(* IEC 61131-3 sources: plc-vscode/tests/st/test-ready/trust-platform/libraries/oscat/oop/src, 12 files *)

(* ---- component_types.st ---- *)
TYPE ComponentStatus :
STRUCT
    Ready : BOOL;
    Error : BOOL;
    ErrorId : WORD;
    Status : BYTE;
END_STRUCT
END_TYPE

TYPE RealRange :
STRUCT
    Low : REAL;
    High : REAL;
END_STRUCT
END_TYPE

TYPE PidGains :
STRUCT
    Kp : REAL := 1.0;
    Tn : REAL := 1.0;
    Tv : REAL := 1.0;
END_STRUCT
END_TYPE

TYPE PiGains :
STRUCT
    Kp : REAL := 1.0;
    Ki : REAL := 1.0;
END_STRUCT
END_TYPE

TYPE SunPosition :
STRUCT
    Azimuth : REAL;
    Elevation : REAL;
    RefractedElevation : REAL;
END_STRUCT
END_TYPE

TYPE SunTimes :
STRUCT
    SolarNoon : TOD;
    Sunrise : TOD;
    Sunset : TOD;
    Declination : REAL;
END_STRUCT
END_TYPE

TYPE BarGraphSnapshot :
STRUCT
    Low : BOOL;
    Q1 : BOOL;
    Q2 : BOOL;
    Q3 : BOOL;
    Q4 : BOOL;
    Q5 : BOOL;
    Q6 : BOOL;
    High : BOOL;
    Alarm : BOOL;
    Status : BYTE;
END_STRUCT
END_TYPE

VAR_GLOBAL CONSTANT
    ComponentErrorNone : WORD := WORD#16#0000;
    ComponentErrorInvalidConfiguration : WORD := WORD#16#1000;
    ComponentErrorNotReady : WORD := WORD#16#1001;
    ComponentErrorQueueFull : WORD := WORD#16#1002;
    ComponentErrorQueueEmpty : WORD := WORD#16#1003;

    DefaultPidKp : REAL := REAL#1.0;
    DefaultPidTn : REAL := REAL#1.0;
    DefaultPidTv : REAL := REAL#1.0;
    DefaultPidLowLimit : REAL := REAL#-1000.0;
    DefaultPidHighLimit : REAL := REAL#1000.0;
    DefaultPidSupervisionBand : REAL := REAL#0.0;
    DefaultPidOffset : REAL := REAL#0.0;

    DefaultPt1Gain : REAL := REAL#1.0;
    DefaultPt1TimeConstant : TIME := T#1s;
    DefaultPulseHighTime : TIME := T#1s;
    DefaultPulseLowTime : TIME := T#1s;
    DefaultCalendarOffsetMinutes : INT := INT#0;
    MaxDwordFifo16Capacity : UINT := UINT#16;
    MaxDwordStack16Capacity : UINT := UINT#16;
    MaxDwordFifo32Capacity : UINT := UINT#32;
    MaxDwordStack32Capacity : UINT := UINT#32;
END_VAR

(* ---- component_interfaces.st ---- *)
INTERFACE IComponent
    PROPERTY Ready : BOOL
    GET
    END_GET
    END_PROPERTY

    PROPERTY Error : BOOL
    GET
    END_GET
    END_PROPERTY

    PROPERTY ErrorId : WORD
    GET
    END_GET
    END_PROPERTY

    PROPERTY Status : BYTE
    GET
    END_GET
    END_PROPERTY

    METHOD Initialize
    END_METHOD

    METHOD Reset
    END_METHOD

    METHOD ClearError
    END_METHOD

    METHOD Snapshot : ComponentStatus
    END_METHOD
END_INTERFACE

INTERFACE IAutomationContext EXTENDS IComponent
    PROPERTY ConstantsLoaded : BOOL
    GET
    END_GET
    END_PROPERTY

    PROPERTY Version : DWORD
    GET
    END_GET
    END_PROPERTY

    PROPERTY Math : CONSTANTS_MATH
    GET
    END_GET
    END_PROPERTY

    PROPERTY Pi2 : REAL
    GET
    END_GET
    END_PROPERTY

    PROPERTY Phys : CONSTANTS_PHYS
    GET
    END_GET
    END_PROPERTY

    PROPERTY LanguageValues : CONSTANTS_LANGUAGE
    GET
    END_GET
    END_PROPERTY

    PROPERTY DefaultLanguage : INT
    GET
    END_GET
    END_PROPERTY

    METHOD LoadConstants : BOOL
    END_METHOD

    METHOD SetDefaultLanguage
    VAR_INPUT
        LanguageIndex : INT;
    END_VAR
    END_METHOD

    METHOD DirectionName : STRING[3]
    VAR_INPUT
        Degrees : REAL;
    END_VAR
    END_METHOD

    METHOD DirectionDegrees : INT
    VAR_INPUT
        Name : STRING[3];
    END_VAR
    END_METHOD
END_INTERFACE

INTERFACE IUnitConverter EXTENDS IComponent
    METHOD KelvinFromCelsius : REAL
    VAR_INPUT
        Celsius : REAL;
    END_VAR
    END_METHOD

    METHOD FahrenheitFromCelsius : REAL
    VAR_INPUT
        Celsius : REAL;
    END_VAR
    END_METHOD

    METHOD CelsiusFromKelvin : REAL
    VAR_INPUT
        Kelvin : REAL;
    END_VAR
    END_METHOD

    METHOD CelsiusFromFahrenheit : REAL
    VAR_INPUT
        Fahrenheit : REAL;
    END_VAR
    END_METHOD

    METHOD MetersPerSecondFromKilometersPerHour : REAL
    VAR_INPUT
        Kmh : REAL;
    END_VAR
    END_METHOD

    METHOD KilometersPerHourFromMetersPerSecond : REAL
    VAR_INPUT
        Mps : REAL;
    END_VAR
    END_METHOD

    METHOD BeaufortFromMetersPerSecond : INT
    VAR_INPUT
        Mps : REAL;
    END_VAR
    END_METHOD

    METHOD AngularFrequencyFromHertz : REAL
    VAR_INPUT
        Frequency : REAL;
    END_VAR
    END_METHOD

    METHOD HertzFromAngularFrequency : REAL
    VAR_INPUT
        AngularFrequency : REAL;
    END_VAR
    END_METHOD

    METHOD PeriodFromHertz : TIME
    VAR_INPUT
        Frequency : REAL;
    END_VAR
    END_METHOD

    METHOD HertzFromPeriod : REAL
    VAR_INPUT
        Period : TIME;
    END_VAR
    END_METHOD

    METHOD WattHoursFromJoules : REAL
    VAR_INPUT
        Joule : REAL;
    END_VAR
    END_METHOD

    METHOD JoulesFromWattHours : REAL
    VAR_INPUT
        WattHour : REAL;
    END_VAR
    END_METHOD

    METHOD JoulesFromCalories : REAL
    VAR_INPUT
        Calorie : REAL;
    END_VAR
    END_METHOD

    METHOD CaloriesFromJoules : REAL
    VAR_INPUT
        Joule : REAL;
    END_VAR
    END_METHOD
END_INTERFACE

INTERFACE IPt1Filter EXTENDS IComponent
    PROPERTY Output : REAL
    GET
    END_GET
    END_PROPERTY

    PROPERTY TimeConstant : TIME
    GET
    END_GET
    END_PROPERTY

    PROPERTY Gain : REAL
    GET
    END_GET
    END_PROPERTY

    METHOD Configure
    VAR_INPUT
        TimeConstant : TIME;
        Gain : REAL;
    END_VAR
    END_METHOD

    METHOD Update : REAL
    VAR_INPUT
        Sample : REAL;
    END_VAR
    END_METHOD
END_INTERFACE

INTERFACE IClosedLoopController EXTENDS IComponent
    PROPERTY Actual : REAL
    GET
    END_GET
    END_PROPERTY

    PROPERTY TargetValue : REAL
    GET
    END_GET
    END_PROPERTY

    PROPERTY Output : REAL
    GET
    END_GET
    END_PROPERTY

    PROPERTY ControlError : REAL
    GET
    END_GET
    END_PROPERTY

    PROPERTY Limited : BOOL
    GET
    END_GET
    END_PROPERTY

    METHOD Update : REAL
    VAR_INPUT
        Actual : REAL;
        Target : REAL;
    END_VAR
    END_METHOD
END_INTERFACE

INTERFACE IPidController EXTENDS IClosedLoopController
    PROPERTY SupervisionBand : REAL
    GET
    END_GET
    END_PROPERTY

    PROPERTY Manual : BOOL
    GET
    END_GET
    END_PROPERTY

    PROPERTY ManualInput : REAL
    GET
    END_GET
    END_PROPERTY

    PROPERTY Offset : REAL
    GET
    END_GET
    END_PROPERTY

    PROPERTY LowLimit : REAL
    GET
    END_GET
    END_PROPERTY

    PROPERTY HighLimit : REAL
    GET
    END_GET
    END_PROPERTY

    PROPERTY Kp : REAL
    GET
    END_GET
    END_PROPERTY

    PROPERTY Tn : REAL
    GET
    END_GET
    END_PROPERTY

    PROPERTY Tv : REAL
    GET
    END_GET
    END_PROPERTY

    METHOD SetKp
    VAR_INPUT
        Kp : REAL;
    END_VAR
    END_METHOD

    METHOD SetIntegralTime
    VAR_INPUT
        Tn : REAL;
    END_VAR
    END_METHOD

    METHOD SetDerivativeTime
    VAR_INPUT
        Tv : REAL;
    END_VAR
    END_METHOD

    METHOD SetSupervisionBand
    VAR_INPUT
        SupervisionBand : REAL;
    END_VAR
    END_METHOD

    METHOD SetOffset
    VAR_INPUT
        Offset : REAL;
    END_VAR
    END_METHOD

    METHOD SetLimits
    VAR_INPUT
        Limits : RealRange;
    END_VAR
    END_METHOD

    METHOD SetManual
    VAR_INPUT
        Manual : BOOL;
        ManualInput : REAL;
    END_VAR
    END_METHOD

    METHOD ApplyGains
    VAR_INPUT
        Gains : PidGains;
    END_VAR
    END_METHOD

    METHOD Configure
    VAR_INPUT
        Gains : PidGains;
        Limits : RealRange;
        SupervisionBand : REAL;
        Offset : REAL;
    END_VAR
    END_METHOD

END_INTERFACE

INTERFACE IHysteresisSwitch EXTENDS IComponent
    PROPERTY MeasuredValue : REAL
    GET
    END_GET
    END_PROPERTY

    PROPERTY LowLimit : REAL
    GET
    END_GET
    END_PROPERTY

    PROPERTY HighLimit : REAL
    GET
    END_GET
    END_PROPERTY

    PROPERTY Q : BOOL
    GET
    END_GET
    END_PROPERTY

    PROPERTY Window : BOOL
    GET
    END_GET
    END_PROPERTY

    METHOD SetLimits
    VAR_INPUT
        Limits : RealRange;
    END_VAR
    END_METHOD

    METHOD Update : BOOL
    VAR_INPUT
        MeasuredValue : REAL;
    END_VAR
    END_METHOD
END_INTERFACE

INTERFACE IPulseGenerator EXTENDS IComponent
    PROPERTY Enabled : BOOL
    GET
    END_GET
    END_PROPERTY

    PROPERTY Output : BOOL
    GET
    END_GET
    END_PROPERTY

    PROPERTY HighTime : TIME
    GET
    END_GET
    END_PROPERTY

    PROPERTY LowTime : TIME
    GET
    END_GET
    END_PROPERTY

    METHOD Configure
    VAR_INPUT
        HighTime : TIME;
        LowTime : TIME;
    END_VAR
    END_METHOD

    METHOD SetEnabled
    VAR_INPUT
        Enabled : BOOL;
    END_VAR
    END_METHOD

    METHOD Update : BOOL
    END_METHOD
END_INTERFACE

INTERFACE IDwordQueue EXTENDS IComponent
    PROPERTY Empty : BOOL
    GET
    END_GET
    END_PROPERTY

    PROPERTY Full : BOOL
    GET
    END_GET
    END_PROPERTY

    PROPERTY Value : DWORD
    GET
    END_GET
    END_PROPERTY

    PROPERTY Capacity : UINT
    GET
    END_GET
    END_PROPERTY

    METHOD Push : BOOL
    VAR_INPUT
        Value : DWORD;
    END_VAR
    END_METHOD

    METHOD TryPop : BOOL
    END_METHOD
END_INTERFACE

INTERFACE IDwordStack EXTENDS IComponent
    PROPERTY Empty : BOOL
    GET
    END_GET
    END_PROPERTY

    PROPERTY Full : BOOL
    GET
    END_GET
    END_PROPERTY

    PROPERTY Value : DWORD
    GET
    END_GET
    END_PROPERTY

    PROPERTY Capacity : UINT
    GET
    END_GET
    END_PROPERTY

    METHOD Push : BOOL
    VAR_INPUT
        Value : DWORD;
    END_VAR
    END_METHOD

    METHOD TryPop : BOOL
    END_METHOD
END_INTERFACE

INTERFACE ICalendarClock EXTENDS IComponent
    PROPERTY Utc : DT
    GET
    END_GET
    END_PROPERTY

    PROPERTY LocalDateTime : DT
    GET
    END_GET
    END_PROPERTY

    PROPERTY LocalDate : DATE
    GET
    END_GET
    END_PROPERTY

    PROPERTY LocalTimeOfDay : TOD
    GET
    END_GET
    END_PROPERTY

    PROPERTY Year : INT
    GET
    END_GET
    END_PROPERTY

    PROPERTY Month : INT
    GET
    END_GET
    END_PROPERTY

    PROPERTY Day : INT
    GET
    END_GET
    END_PROPERTY

    PROPERTY Weekday : INT
    GET
    END_GET
    END_PROPERTY

    PROPERTY OffsetMinutes : INT
    GET
    END_GET
    END_PROPERTY

    PROPERTY DstEnabled : BOOL
    GET
    END_GET
    END_PROPERTY

    PROPERTY DstOn : BOOL
    GET
    END_GET
    END_PROPERTY

    PROPERTY LanguageIndex : INT
    GET
    END_GET
    END_PROPERTY

    PROPERTY Longitude : REAL
    GET
    END_GET
    END_PROPERTY

    PROPERTY Latitude : REAL
    GET
    END_GET
    END_PROPERTY

    PROPERTY Sunrise : TOD
    GET
    END_GET
    END_PROPERTY

    PROPERTY Sunset : TOD
    GET
    END_GET
    END_PROPERTY

    PROPERTY SolarNoon : TOD
    GET
    END_GET
    END_PROPERTY

    PROPERTY SolarElevation : REAL
    GET
    END_GET
    END_PROPERTY

    PROPERTY SolarHorizontalProjection : REAL
    GET
    END_GET
    END_PROPERTY

    PROPERTY SolarVerticalProjection : REAL
    GET
    END_GET
    END_PROPERTY

    PROPERTY Night : BOOL
    GET
    END_GET
    END_PROPERTY

    PROPERTY Holiday : BOOL
    GET
    END_GET
    END_PROPERTY

    PROPERTY HolidayName : STRING[30]
    GET
    END_GET
    END_PROPERTY

    PROPERTY WorkWeek : INT
    GET
    END_GET
    END_PROPERTY

    METHOD Configure
    VAR_INPUT
        LocationLatitude : REAL;
        LocationLongitude : REAL;
        OffsetMinutes : INT;
        DstEnabled : BOOL;
        LanguageIndex : INT;
    END_VAR
    END_METHOD

    METHOD Update
    VAR_INPUT
        Utc : DT;
    END_VAR
    END_METHOD

    METHOD CalculateSunPosition : SunPosition
    VAR_INPUT
        Utc : DT;
        Latitude : REAL;
        Longitude : REAL;
    END_VAR
    END_METHOD

    METHOD CalculateSunTime : SunTimes
    VAR_INPUT
        UtcDate : DATE;
        Latitude : REAL;
        Longitude : REAL;
        Horizon : REAL;
    END_VAR
    END_METHOD
END_INTERFACE

(* ---- automation_context.st ---- *)
FUNCTION_BLOCK AutomationContext IMPLEMENTS IAutomationContext
VAR
    ReadyValue : BOOL;
    ErrorValue : BOOL;
    ErrorIdValue : WORD;
    StatusValue : BYTE;
    ConstantsLoadedValue : BOOL;
END_VAR

METHOD PUBLIC Initialize
ApplyConstantsLoadResult(Loaded := OSCAT_BASIC_Constants());
END_METHOD

METHOD PUBLIC Reset
ClearError();
ConstantsLoadedValue := FALSE;
END_METHOD

METHOD PUBLIC ClearError
ErrorValue := FALSE;
ErrorIdValue := ComponentErrorNone;
StatusValue := BYTE#0;
END_METHOD

METHOD PUBLIC Snapshot : ComponentStatus
VAR
    Result : ComponentStatus;
END_VAR
Result.Ready := ReadyValue;
Result.Error := ErrorValue;
Result.ErrorId := ErrorIdValue;
Result.Status := StatusValue;
Snapshot := Result;
END_METHOD

METHOD PUBLIC LoadConstants : BOOL
LoadConstants := OSCAT_BASIC_Constants();
ApplyConstantsLoadResult(Loaded := LoadConstants);
END_METHOD

METHOD PRIVATE ApplyConstantsLoadResult
VAR_INPUT
    Loaded : BOOL;
END_VAR
ConstantsLoadedValue := Loaded;
ReadyValue := Loaded;
IF Loaded THEN
    ClearError();
ELSE
    ErrorValue := TRUE;
    ErrorIdValue := ComponentErrorNotReady;
    StatusValue := BYTE#1;
END_IF;
END_METHOD

METHOD PUBLIC SetDefaultLanguage
VAR_INPUT
    LanguageIndex : INT;
END_VAR
IF NOT ConstantsLoadedValue AND NOT LoadConstants() THEN
    ErrorValue := TRUE;
    ErrorIdValue := ComponentErrorNotReady;
    StatusValue := BYTE#1;
ELSIF LanguageIndex >= INT#1 AND LanguageIndex <= LANGUAGE.LMAX THEN
    LANGUAGE.DEFAULT := LanguageIndex;
    ClearError();
ELSE
    ErrorValue := TRUE;
    ErrorIdValue := ComponentErrorInvalidConfiguration;
    StatusValue := BYTE#1;
END_IF;
END_METHOD

METHOD PUBLIC DirectionName : STRING[3]
VAR_INPUT
    Degrees : REAL;
END_VAR
IF NOT ConstantsLoadedValue AND NOT LoadConstants() THEN
    DirectionName := '';
ELSE
    DirectionName := DEG_TO_DIR(DEG := REAL_TO_INT(Degrees), N := INT#4, L := LANGUAGE.DEFAULT);
END_IF;
END_METHOD

METHOD PUBLIC DirectionDegrees : INT
VAR_INPUT
    Name : STRING[3];
END_VAR
IF NOT ConstantsLoadedValue AND NOT LoadConstants() THEN
    DirectionDegrees := INT#0;
ELSE
    DirectionDegrees := DIR_TO_DEG(DIR := Name, L := LANGUAGE.DEFAULT);
END_IF;
END_METHOD

PUBLIC PROPERTY Ready : BOOL
GET
    Ready := ReadyValue;
END_GET
END_PROPERTY

PUBLIC PROPERTY Error : BOOL
GET
    Error := ErrorValue;
END_GET
END_PROPERTY

PUBLIC PROPERTY ErrorId : WORD
GET
    ErrorId := ErrorIdValue;
END_GET
END_PROPERTY

PUBLIC PROPERTY Status : BYTE
GET
    Status := StatusValue;
END_GET
END_PROPERTY

PUBLIC PROPERTY ConstantsLoaded : BOOL
GET
    ConstantsLoaded := ConstantsLoadedValue OR g_oscat_constants_loaded;
END_GET
END_PROPERTY

PUBLIC PROPERTY Version : DWORD
GET
    Version := OSCAT_VERSION(IN := FALSE);
END_GET
END_PROPERTY

PUBLIC PROPERTY Math : CONSTANTS_MATH
GET
    Math := MATH;
END_GET
END_PROPERTY

PUBLIC PROPERTY Pi2 : REAL
GET
    Pi2 := MATH.PI2;
END_GET
END_PROPERTY

PUBLIC PROPERTY Phys : CONSTANTS_PHYS
GET
    Phys := PHYS;
END_GET
END_PROPERTY

PUBLIC PROPERTY LanguageValues : CONSTANTS_LANGUAGE
GET
    LanguageValues := LANGUAGE;
END_GET
END_PROPERTY

PUBLIC PROPERTY DefaultLanguage : INT
GET
    DefaultLanguage := LANGUAGE.DEFAULT;
END_GET
END_PROPERTY
END_FUNCTION_BLOCK

(* ---- calendar.st ---- *)
FUNCTION_BLOCK CalendarClock IMPLEMENTS ICalendarClock
VAR
    ReadyValue : BOOL;
    ErrorValue : BOOL;
    ErrorIdValue : WORD;
    StatusValue : BYTE;
    CalendarData : CALENDAR;
    Holidays : ARRAY[0..29] OF HOLIDAY_DATA;
    CalendarFb : CALENDAR_CALC;
    SunPositionFb : SUN_POS;
    SunTimeFb : SUN_TIME;
END_VAR

METHOD PUBLIC Initialize
ReadyValue := TRUE;
OSCAT_BASIC_Constants();
CalendarData.OFFSET := DefaultCalendarOffsetMinutes;
CalendarData.LANGUAGE := LANGUAGE.DEFAULT;
ClearError();
END_METHOD

METHOD PUBLIC Reset
ClearError();
END_METHOD

METHOD PUBLIC ClearError
ErrorValue := FALSE;
ErrorIdValue := ComponentErrorNone;
StatusValue := BYTE#0;
END_METHOD

METHOD PUBLIC Snapshot : ComponentStatus
VAR
    Result : ComponentStatus;
END_VAR
Result.Ready := ReadyValue;
Result.Error := ErrorValue;
Result.ErrorId := ErrorIdValue;
Result.Status := StatusValue;
Snapshot := Result;
END_METHOD

METHOD PUBLIC Configure
VAR_INPUT
    LocationLatitude : REAL;
    LocationLongitude : REAL;
    OffsetMinutes : INT;
    DstEnabled : BOOL;
    LanguageIndex : INT;
END_VAR
IF NOT ReadyValue THEN
    Initialize();
END_IF;
CalendarData.LATITUDE := LocationLatitude;
CalendarData.LONGITUDE := LocationLongitude;
CalendarData.OFFSET := OffsetMinutes;
CalendarData.DST_EN := DstEnabled;
CalendarData.LANGUAGE := LanguageIndex;
ClearError();
END_METHOD

METHOD PUBLIC Update
VAR_INPUT
    Utc : DT;
END_VAR
IF NOT ReadyValue THEN
    Initialize();
END_IF;
CalendarData.UTC := Utc;
CalendarFb(SPE := TRUE, H := REAL#-0.8333333, XCAL := CalendarData, HOLIDAYS := Holidays);
END_METHOD

METHOD PUBLIC CalculateSunPosition : SunPosition
VAR_INPUT
    Utc : DT;
    Latitude : REAL;
    Longitude : REAL;
END_VAR
VAR
    Result : SunPosition;
END_VAR
OSCAT_BASIC_Constants();
SunPositionFb(LATITUDE := Latitude, LONGITUDE := Longitude, UTC := Utc);
Result.Azimuth := SunPositionFb.B;
Result.Elevation := SunPositionFb.H;
Result.RefractedElevation := SunPositionFb.HR;
CalculateSunPosition := Result;
END_METHOD

METHOD PUBLIC CalculateSunTime : SunTimes
VAR_INPUT
    UtcDate : DATE;
    Latitude : REAL;
    Longitude : REAL;
    Horizon : REAL;
END_VAR
VAR
    Result : SunTimes;
END_VAR
OSCAT_BASIC_Constants();
SunTimeFb(LATITUDE := Latitude, LONGITUDE := Longitude, UTC := UtcDate, H := Horizon);
Result.SolarNoon := SunTimeFb.MIDDAY;
Result.Sunrise := SunTimeFb.SUN_RISE;
Result.Sunset := SunTimeFb.SUN_SET;
Result.Declination := SunTimeFb.SUN_DECLINATION;
CalculateSunTime := Result;
END_METHOD

PUBLIC PROPERTY Ready : BOOL
GET
    Ready := ReadyValue;
END_GET
END_PROPERTY

PUBLIC PROPERTY Error : BOOL
GET
    Error := ErrorValue;
END_GET
END_PROPERTY

PUBLIC PROPERTY ErrorId : WORD
GET
    ErrorId := ErrorIdValue;
END_GET
END_PROPERTY

PUBLIC PROPERTY Status : BYTE
GET
    Status := StatusValue;
END_GET
END_PROPERTY

PUBLIC PROPERTY Utc : DT
GET
    Utc := CalendarData.UTC;
END_GET
END_PROPERTY

PUBLIC PROPERTY LocalDateTime : DT
GET
    LocalDateTime := CalendarData.LOCAL_DT;
END_GET
END_PROPERTY

PUBLIC PROPERTY LocalDate : DATE
GET
    LocalDate := CalendarData.LOCAL_DATE;
END_GET
END_PROPERTY

PUBLIC PROPERTY LocalTimeOfDay : TOD
GET
    LocalTimeOfDay := CalendarData.LOCAL_TOD;
END_GET
END_PROPERTY

PUBLIC PROPERTY Year : INT
GET
    Year := CalendarData.YEAR;
END_GET
END_PROPERTY

PUBLIC PROPERTY Month : INT
GET
    Month := CalendarData.MONTH;
END_GET
END_PROPERTY

PUBLIC PROPERTY Day : INT
GET
    Day := CalendarData.DAY;
END_GET
END_PROPERTY

PUBLIC PROPERTY Weekday : INT
GET
    Weekday := CalendarData.WEEKDAY;
END_GET
END_PROPERTY

PUBLIC PROPERTY OffsetMinutes : INT
GET
    OffsetMinutes := CalendarData.OFFSET;
END_GET
END_PROPERTY

PUBLIC PROPERTY DstEnabled : BOOL
GET
    DstEnabled := CalendarData.DST_EN;
END_GET
END_PROPERTY

PUBLIC PROPERTY DstOn : BOOL
GET
    DstOn := CalendarData.DST_ON;
END_GET
END_PROPERTY

PUBLIC PROPERTY LanguageIndex : INT
GET
    LanguageIndex := CalendarData.LANGUAGE;
END_GET
END_PROPERTY

PUBLIC PROPERTY Longitude : REAL
GET
    Longitude := CalendarData.LONGITUDE;
END_GET
END_PROPERTY

PUBLIC PROPERTY Latitude : REAL
GET
    Latitude := CalendarData.LATITUDE;
END_GET
END_PROPERTY

PUBLIC PROPERTY Sunrise : TOD
GET
    Sunrise := CalendarData.SUN_RISE;
END_GET
END_PROPERTY

PUBLIC PROPERTY Sunset : TOD
GET
    Sunset := CalendarData.SUN_SET;
END_GET
END_PROPERTY

PUBLIC PROPERTY SolarNoon : TOD
GET
    SolarNoon := CalendarData.SUN_MIDDAY;
END_GET
END_PROPERTY

PUBLIC PROPERTY SolarElevation : REAL
GET
    (* OSCAT classic keeps the historical SUN_HEIGTH spelling. *)
    SolarElevation := CalendarData.SUN_HEIGTH;
END_GET
END_PROPERTY

PUBLIC PROPERTY SolarHorizontalProjection : REAL
GET
    SolarHorizontalProjection := CalendarData.SUN_HOR;
END_GET
END_PROPERTY

PUBLIC PROPERTY SolarVerticalProjection : REAL
GET
    SolarVerticalProjection := CalendarData.SUN_VER;
END_GET
END_PROPERTY

PUBLIC PROPERTY Night : BOOL
GET
    Night := CalendarData.NIGHT;
END_GET
END_PROPERTY

PUBLIC PROPERTY Holiday : BOOL
GET
    Holiday := CalendarData.HOLIDAY;
END_GET
END_PROPERTY

PUBLIC PROPERTY HolidayName : STRING[30]
GET
    HolidayName := CalendarData.HOLY_NAME;
END_GET
END_PROPERTY

PUBLIC PROPERTY WorkWeek : INT
GET
    WorkWeek := CalendarData.WORK_WEEK;
END_GET
END_PROPERTY
END_FUNCTION_BLOCK

FUNCTION_BLOCK HolidayCalendar IMPLEMENTS IComponent
VAR
    ReadyValue : BOOL;
    ErrorValue : BOOL;
    ErrorIdValue : WORD;
    StatusValue : BYTE;
    HolidayValue : BOOL;
    NameValue : STRING[30];
    LanguageIndexValue : INT := INT#1;
    FridayAsHolidayValue : BOOL;
    SaturdayAsHolidayValue : BOOL;
    SundayAsHolidayValue : BOOL;
    Holidays : ARRAY[0..29] OF HOLIDAY_DATA;
    HolidayFb : HOLIDAY;
END_VAR

METHOD PUBLIC Initialize
ReadyValue := TRUE;
OSCAT_BASIC_Constants();
ClearError();
END_METHOD

METHOD PUBLIC Reset
HolidayValue := FALSE;
NameValue := '';
ClearError();
END_METHOD

METHOD PUBLIC ClearError
ErrorValue := FALSE;
ErrorIdValue := ComponentErrorNone;
StatusValue := BYTE#0;
END_METHOD

METHOD PUBLIC Snapshot : ComponentStatus
VAR
    Result : ComponentStatus;
END_VAR
Result.Ready := ReadyValue;
Result.Error := ErrorValue;
Result.ErrorId := ErrorIdValue;
Result.Status := StatusValue;
Snapshot := Result;
END_METHOD

METHOD PUBLIC Configure
VAR_INPUT
    LanguageIndex : INT;
    FridayAsHoliday : BOOL;
    SaturdayAsHoliday : BOOL;
    SundayAsHoliday : BOOL;
END_VAR
LanguageIndexValue := LanguageIndex;
FridayAsHolidayValue := FridayAsHoliday;
SaturdayAsHolidayValue := SaturdayAsHoliday;
SundayAsHolidayValue := SundayAsHoliday;
ClearError();
END_METHOD

METHOD PUBLIC SetHoliday
VAR_INPUT
    Index : INT;
    Month : SINT;
    Day : SINT;
    Use : SINT;
    Name : STRING[30];
END_VAR
IF Index < INT#0 OR Index > INT#29 THEN
    ErrorValue := TRUE;
    ErrorIdValue := ComponentErrorInvalidConfiguration;
    StatusValue := BYTE#1;
ELSE
    Holidays[Index].MONTH := Month;
    Holidays[Index].DAY := Day;
    Holidays[Index].USE := Use;
    Holidays[Index].NAME := Name;
    ClearError();
END_IF;
END_METHOD

METHOD PUBLIC Update : BOOL
VAR_INPUT
    DateIn : DATE;
END_VAR
HolidayFb(
    DATE_IN := DateIn,
    LANGU := LanguageIndexValue,
    FRIDAY := FridayAsHolidayValue,
    SATURDAY := SaturdayAsHolidayValue,
    SUNDAY := SundayAsHolidayValue,
    HOLIDAYS := Holidays
);
HolidayValue := HolidayFb.Y;
NameValue := HolidayFb.NAME;
Update := HolidayValue;
END_METHOD

PUBLIC PROPERTY Ready : BOOL
GET
    Ready := ReadyValue;
END_GET
END_PROPERTY

PUBLIC PROPERTY Error : BOOL
GET
    Error := ErrorValue;
END_GET
END_PROPERTY

PUBLIC PROPERTY ErrorId : WORD
GET
    ErrorId := ErrorIdValue;
END_GET
END_PROPERTY

PUBLIC PROPERTY Status : BYTE
GET
    Status := StatusValue;
END_GET
END_PROPERTY

PUBLIC PROPERTY Holiday : BOOL
GET
    Holiday := HolidayValue;
END_GET
END_PROPERTY

PUBLIC PROPERTY Name : STRING[30]
GET
    Name := NameValue;
END_GET
END_PROPERTY
END_FUNCTION_BLOCK

FUNCTION_BLOCK RtcClock IMPLEMENTS IComponent
VAR
    ReadyValue : BOOL;
    ErrorValue : BOOL;
    ErrorIdValue : WORD;
    StatusValue : BYTE;
    UtcDateTimeValue : DT;
    LocalDateTimeValue : DT;
    DstOnValue : BOOL;
    MillisecondsValue : INT;
    DstEnabledValue : BOOL;
    OffsetMinutesValue : INT;
    RtcFb : RTC_2;
END_VAR

METHOD PUBLIC Initialize
ReadyValue := TRUE;
ClearError();
END_METHOD

METHOD PUBLIC Reset
UtcDateTimeValue := DT#1970-01-01-00:00:00;
LocalDateTimeValue := DT#1970-01-01-00:00:00;
MillisecondsValue := INT#0;
ClearError();
END_METHOD

METHOD PUBLIC ClearError
ErrorValue := FALSE;
ErrorIdValue := ComponentErrorNone;
StatusValue := BYTE#0;
END_METHOD

METHOD PUBLIC Snapshot : ComponentStatus
VAR
    Result : ComponentStatus;
END_VAR
Result.Ready := ReadyValue;
Result.Error := ErrorValue;
Result.ErrorId := ErrorIdValue;
Result.Status := StatusValue;
Snapshot := Result;
END_METHOD

METHOD PUBLIC SetClock
VAR_INPUT
    InitialDateTime : DT;
    Milliseconds : INT;
    DstEnabled : BOOL;
    OffsetMinutes : INT;
END_VAR
DstEnabledValue := DstEnabled;
OffsetMinutesValue := OffsetMinutes;
RtcFb(SET_RTC := TRUE, SDT := InitialDateTime, SMS := Milliseconds, DEN := DstEnabledValue, OFS := OffsetMinutesValue);
UtcDateTimeValue := RtcFb.UDT;
LocalDateTimeValue := RtcFb.LOCAL_DT;
DstOnValue := RtcFb.DSO;
MillisecondsValue := RtcFb.XMS;
ClearError();
END_METHOD

METHOD PUBLIC Update
RtcFb(SET_RTC := FALSE, SDT := UtcDateTimeValue, SMS := MillisecondsValue, DEN := DstEnabledValue, OFS := OffsetMinutesValue);
UtcDateTimeValue := RtcFb.UDT;
LocalDateTimeValue := RtcFb.LOCAL_DT;
DstOnValue := RtcFb.DSO;
MillisecondsValue := RtcFb.XMS;
END_METHOD

PUBLIC PROPERTY Ready : BOOL
GET
    Ready := ReadyValue;
END_GET
END_PROPERTY

PUBLIC PROPERTY Error : BOOL
GET
    Error := ErrorValue;
END_GET
END_PROPERTY

PUBLIC PROPERTY ErrorId : WORD
GET
    ErrorId := ErrorIdValue;
END_GET
END_PROPERTY

PUBLIC PROPERTY Status : BYTE
GET
    Status := StatusValue;
END_GET
END_PROPERTY

PUBLIC PROPERTY UtcDateTime : DT
GET
    UtcDateTime := UtcDateTimeValue;
END_GET
END_PROPERTY

PUBLIC PROPERTY LocalDateTime : DT
GET
    LocalDateTime := LocalDateTimeValue;
END_GET
END_PROPERTY

PUBLIC PROPERTY DstOn : BOOL
GET
    DstOn := DstOnValue;
END_GET
END_PROPERTY

PUBLIC PROPERTY Milliseconds : INT
GET
    Milliseconds := MillisecondsValue;
END_GET
END_PROPERTY
END_FUNCTION_BLOCK

(* ---- control.st ---- *)
FUNCTION_BLOCK PidController IMPLEMENTS IPidController
VAR
    ReadyValue : BOOL;
    ErrorValue : BOOL;
    ErrorIdValue : WORD;
    StatusValue : BYTE;
    ActualValue : REAL;
    SetpointValue : REAL;
    SupervisionBandValue : REAL := DefaultPidSupervisionBand;
    ManualValue : BOOL;
    ManualInputValue : REAL;
    OffsetValue : REAL := DefaultPidOffset;
    OutputValue : REAL;
    ControlErrorValue : REAL;
    LimitedValue : BOOL;
    LowLimitValue : REAL := DefaultPidLowLimit;
    HighLimitValue : REAL := DefaultPidHighLimit;
    KpValue : REAL := DefaultPidKp;
    TnValue : REAL := DefaultPidTn;
    TvValue : REAL := DefaultPidTv;
    ResetRequested : BOOL;
    ControllerFb : CTRL_PID;
END_VAR

METHOD PUBLIC Initialize
ReadyValue := TRUE;
ClearError();
END_METHOD

METHOD PUBLIC Reset
ResetRequested := TRUE;
OutputValue := REAL#0.0;
ControlErrorValue := REAL#0.0;
LimitedValue := FALSE;
ClearError();
END_METHOD

METHOD PUBLIC ClearError
ErrorValue := FALSE;
ErrorIdValue := ComponentErrorNone;
StatusValue := BYTE#0;
END_METHOD

METHOD PUBLIC Snapshot : ComponentStatus
VAR
    Result : ComponentStatus;
END_VAR
Result.Ready := ReadyValue;
Result.Error := ErrorValue;
Result.ErrorId := ErrorIdValue;
Result.Status := StatusValue;
Snapshot := Result;
END_METHOD

METHOD PUBLIC SetKp
VAR_INPUT
    Kp : REAL;
END_VAR
KpValue := Kp;
ClearError();
END_METHOD

METHOD PUBLIC SetIntegralTime
VAR_INPUT
    Tn : REAL;
END_VAR
TnValue := Tn;
ClearError();
END_METHOD

METHOD PUBLIC SetDerivativeTime
VAR_INPUT
    Tv : REAL;
END_VAR
TvValue := Tv;
ClearError();
END_METHOD

METHOD PUBLIC SetSupervisionBand
VAR_INPUT
    SupervisionBand : REAL;
END_VAR
SupervisionBandValue := SupervisionBand;
ClearError();
END_METHOD

METHOD PUBLIC SetOffset
VAR_INPUT
    Offset : REAL;
END_VAR
OffsetValue := Offset;
ClearError();
END_METHOD

METHOD PUBLIC SetLimits
VAR_INPUT
    Limits : RealRange;
END_VAR
IF Limits.High < Limits.Low THEN
    ErrorValue := TRUE;
    ErrorIdValue := ComponentErrorInvalidConfiguration;
    StatusValue := BYTE#1;
ELSE
    LowLimitValue := Limits.Low;
    HighLimitValue := Limits.High;
    ClearError();
END_IF;
END_METHOD

METHOD PUBLIC SetManual
VAR_INPUT
    Manual : BOOL;
    ManualInput : REAL;
END_VAR
ManualValue := Manual;
ManualInputValue := ManualInput;
ClearError();
END_METHOD

METHOD PUBLIC ApplyGains
VAR_INPUT
    Gains : PidGains;
END_VAR
KpValue := Gains.Kp;
TnValue := Gains.Tn;
TvValue := Gains.Tv;
ClearError();
END_METHOD

METHOD PUBLIC Configure
VAR_INPUT
    Gains : PidGains;
    Limits : RealRange;
    SupervisionBand : REAL;
    Offset : REAL;
END_VAR
IF Limits.High < Limits.Low THEN
    ErrorValue := TRUE;
    ErrorIdValue := ComponentErrorInvalidConfiguration;
    StatusValue := BYTE#1;
ELSE
    KpValue := Gains.Kp;
    TnValue := Gains.Tn;
    TvValue := Gains.Tv;
    LowLimitValue := Limits.Low;
    HighLimitValue := Limits.High;
    SupervisionBandValue := SupervisionBand;
    OffsetValue := Offset;
    ClearError();
END_IF;
END_METHOD

METHOD PUBLIC Update : REAL
VAR_INPUT
    Actual : REAL;
    Target : REAL;
END_VAR
IF NOT ReadyValue THEN
    ReadyValue := TRUE;
END_IF;
ActualValue := Actual;
SetpointValue := Target;
ControllerFb(
    ACT := ActualValue,
    SET_POINT := SetpointValue,
    SUP := SupervisionBandValue,
    OFS := OffsetValue,
    M_I := ManualInputValue,
    MAN := ManualValue,
    RST := ResetRequested,
    KP := KpValue,
    TN := TnValue,
    TV := TvValue,
    LL := LowLimitValue,
    LH := HighLimitValue
);
ResetRequested := FALSE;
OutputValue := ControllerFb.Y;
ControlErrorValue := ControllerFb.DIFF;
LimitedValue := ControllerFb.LIM;
Update := OutputValue;
END_METHOD

PUBLIC PROPERTY Ready : BOOL
GET
    Ready := ReadyValue;
END_GET
END_PROPERTY

PUBLIC PROPERTY Error : BOOL
GET
    Error := ErrorValue;
END_GET
END_PROPERTY

PUBLIC PROPERTY ErrorId : WORD
GET
    ErrorId := ErrorIdValue;
END_GET
END_PROPERTY

PUBLIC PROPERTY Status : BYTE
GET
    Status := StatusValue;
END_GET
END_PROPERTY

PUBLIC PROPERTY Actual : REAL
GET
    Actual := ActualValue;
END_GET
END_PROPERTY

PUBLIC PROPERTY TargetValue : REAL
GET
    TargetValue := SetpointValue;
END_GET
END_PROPERTY

PUBLIC PROPERTY SupervisionBand : REAL
GET
    SupervisionBand := SupervisionBandValue;
END_GET
END_PROPERTY

PUBLIC PROPERTY Manual : BOOL
GET
    Manual := ManualValue;
END_GET
END_PROPERTY

PUBLIC PROPERTY ManualInput : REAL
GET
    ManualInput := ManualInputValue;
END_GET
END_PROPERTY

PUBLIC PROPERTY Offset : REAL
GET
    Offset := OffsetValue;
END_GET
END_PROPERTY

PUBLIC PROPERTY Output : REAL
GET
    Output := OutputValue;
END_GET
END_PROPERTY

PUBLIC PROPERTY ControlError : REAL
GET
    ControlError := ControlErrorValue;
END_GET
END_PROPERTY

PUBLIC PROPERTY Limited : BOOL
GET
    Limited := LimitedValue;
END_GET
END_PROPERTY

PUBLIC PROPERTY LowLimit : REAL
GET
    LowLimit := LowLimitValue;
END_GET
END_PROPERTY

PUBLIC PROPERTY HighLimit : REAL
GET
    HighLimit := HighLimitValue;
END_GET
END_PROPERTY

PUBLIC PROPERTY Kp : REAL
GET
    Kp := KpValue;
END_GET
END_PROPERTY

PUBLIC PROPERTY Tn : REAL
GET
    Tn := TnValue;
END_GET
END_PROPERTY

PUBLIC PROPERTY Tv : REAL
GET
    Tv := TvValue;
END_GET
END_PROPERTY
END_FUNCTION_BLOCK

FUNCTION_BLOCK PiController IMPLEMENTS IClosedLoopController
VAR
    ReadyValue : BOOL;
    ErrorValue : BOOL;
    ErrorIdValue : WORD;
    StatusValue : BYTE;
    ActualValue : REAL;
    SetpointValue : REAL;
    OutputValue : REAL;
    ControlErrorValue : REAL;
    LimitedValue : BOOL;
    SupervisionBandValue : REAL := DefaultPidSupervisionBand;
    ManualValue : BOOL;
    ManualInputValue : REAL;
    OffsetValue : REAL := DefaultPidOffset;
    LowLimitValue : REAL := DefaultPidLowLimit;
    HighLimitValue : REAL := DefaultPidHighLimit;
    KpValue : REAL := DefaultPidKp;
    KiValue : REAL := REAL#1.0;
    ResetRequested : BOOL;
    ControllerFb : CTRL_PI;
END_VAR

METHOD PUBLIC Initialize
ReadyValue := TRUE;
ClearError();
END_METHOD

METHOD PUBLIC Reset
ResetRequested := TRUE;
OutputValue := REAL#0.0;
ControlErrorValue := REAL#0.0;
LimitedValue := FALSE;
ClearError();
END_METHOD

METHOD PUBLIC ClearError
ErrorValue := FALSE;
ErrorIdValue := ComponentErrorNone;
StatusValue := BYTE#0;
END_METHOD

METHOD PUBLIC Snapshot : ComponentStatus
VAR
    Result : ComponentStatus;
END_VAR
Result.Ready := ReadyValue;
Result.Error := ErrorValue;
Result.ErrorId := ErrorIdValue;
Result.Status := StatusValue;
Snapshot := Result;
END_METHOD

METHOD PUBLIC Configure
VAR_INPUT
    Gains : PiGains;
    Limits : RealRange;
    SupervisionBand : REAL;
    Offset : REAL;
END_VAR
IF Limits.High < Limits.Low THEN
    ErrorValue := TRUE;
    ErrorIdValue := ComponentErrorInvalidConfiguration;
    StatusValue := BYTE#1;
ELSE
    KpValue := Gains.Kp;
    KiValue := Gains.Ki;
    LowLimitValue := Limits.Low;
    HighLimitValue := Limits.High;
    SupervisionBandValue := SupervisionBand;
    OffsetValue := Offset;
    ClearError();
END_IF;
END_METHOD

METHOD PUBLIC SetManual
VAR_INPUT
    Manual : BOOL;
    ManualInput : REAL;
END_VAR
ManualValue := Manual;
ManualInputValue := ManualInput;
ClearError();
END_METHOD

METHOD PUBLIC Update : REAL
VAR_INPUT
    Actual : REAL;
    Target : REAL;
END_VAR
IF NOT ReadyValue THEN
    ReadyValue := TRUE;
END_IF;
ActualValue := Actual;
SetpointValue := Target;
ControllerFb(
    ACT := ActualValue,
    SET_POINT := SetpointValue,
    SUP := SupervisionBandValue,
    OFS := OffsetValue,
    M_I := ManualInputValue,
    MAN := ManualValue,
    RST := ResetRequested,
    KP := KpValue,
    KI := KiValue,
    LL := LowLimitValue,
    LH := HighLimitValue
);
ResetRequested := FALSE;
OutputValue := ControllerFb.Y;
ControlErrorValue := ControllerFb.DIFF;
LimitedValue := ControllerFb.LIM;
Update := OutputValue;
END_METHOD

PUBLIC PROPERTY Ready : BOOL
GET
    Ready := ReadyValue;
END_GET
END_PROPERTY

PUBLIC PROPERTY Error : BOOL
GET
    Error := ErrorValue;
END_GET
END_PROPERTY

PUBLIC PROPERTY ErrorId : WORD
GET
    ErrorId := ErrorIdValue;
END_GET
END_PROPERTY

PUBLIC PROPERTY Status : BYTE
GET
    Status := StatusValue;
END_GET
END_PROPERTY

PUBLIC PROPERTY Actual : REAL
GET
    Actual := ActualValue;
END_GET
END_PROPERTY

PUBLIC PROPERTY TargetValue : REAL
GET
    TargetValue := SetpointValue;
END_GET
END_PROPERTY

PUBLIC PROPERTY Output : REAL
GET
    Output := OutputValue;
END_GET
END_PROPERTY

PUBLIC PROPERTY ControlError : REAL
GET
    ControlError := ControlErrorValue;
END_GET
END_PROPERTY

PUBLIC PROPERTY Limited : BOOL
GET
    Limited := LimitedValue;
END_GET
END_PROPERTY
END_FUNCTION_BLOCK

FUNCTION_BLOCK PwmController IMPLEMENTS IComponent
VAR
    ReadyValue : BOOL;
    ErrorValue : BOOL;
    ErrorIdValue : WORD;
    StatusValue : BYTE;
    OutputValue : BOOL;
    FrequencyValue : REAL;
    ManualValue : BOOL;
    ManualInputValue : REAL;
    ControllerFb : CTRL_PWM;
END_VAR

METHOD PUBLIC Initialize
ReadyValue := TRUE;
ClearError();
END_METHOD

METHOD PUBLIC Reset
ControllerFb(CI := REAL#0.0, MAN_IN := REAL#0.0, MANUAL := FALSE, F := REAL#0.0);
OutputValue := ControllerFb.Q;
ClearError();
END_METHOD

METHOD PUBLIC ClearError
ErrorValue := FALSE;
ErrorIdValue := ComponentErrorNone;
StatusValue := BYTE#0;
END_METHOD

METHOD PUBLIC Snapshot : ComponentStatus
VAR
    Result : ComponentStatus;
END_VAR
Result.Ready := ReadyValue;
Result.Error := ErrorValue;
Result.ErrorId := ErrorIdValue;
Result.Status := StatusValue;
Snapshot := Result;
END_METHOD

METHOD PUBLIC Configure
VAR_INPUT
    Frequency : REAL;
END_VAR
FrequencyValue := Frequency;
ClearError();
END_METHOD

METHOD PUBLIC SetManual
VAR_INPUT
    Manual : BOOL;
    ManualInput : REAL;
END_VAR
ManualValue := Manual;
ManualInputValue := ManualInput;
ClearError();
END_METHOD

METHOD PUBLIC Update : BOOL
VAR_INPUT
    ControlInput : REAL;
END_VAR
IF NOT ReadyValue THEN
    ReadyValue := TRUE;
END_IF;
ControllerFb(CI := ControlInput, MAN_IN := ManualInputValue, MANUAL := ManualValue, F := FrequencyValue);
OutputValue := ControllerFb.Q;
Update := OutputValue;
END_METHOD

PUBLIC PROPERTY Ready : BOOL
GET
    Ready := ReadyValue;
END_GET
END_PROPERTY

PUBLIC PROPERTY Error : BOOL
GET
    Error := ErrorValue;
END_GET
END_PROPERTY

PUBLIC PROPERTY ErrorId : WORD
GET
    ErrorId := ErrorIdValue;
END_GET
END_PROPERTY

PUBLIC PROPERTY Status : BYTE
GET
    Status := StatusValue;
END_GET
END_PROPERTY

PUBLIC PROPERTY Output : BOOL
GET
    Output := OutputValue;
END_GET
END_PROPERTY

PUBLIC PROPERTY Frequency : REAL
GET
    Frequency := FrequencyValue;
END_GET
END_PROPERTY
END_FUNCTION_BLOCK

FUNCTION_BLOCK HysteresisSwitch IMPLEMENTS IHysteresisSwitch
VAR
    ReadyValue : BOOL;
    ErrorValue : BOOL;
    ErrorIdValue : WORD;
    StatusValue : BYTE;
    MeasuredValueValue : REAL;
    LowLimitValue : REAL;
    HighLimitValue : REAL;
    QValue : BOOL;
    WindowValue : BOOL;
END_VAR

METHOD PUBLIC Initialize
ReadyValue := TRUE;
ClearError();
END_METHOD

METHOD PUBLIC Reset
QValue := FALSE;
WindowValue := FALSE;
ClearError();
END_METHOD

METHOD PUBLIC ClearError
ErrorValue := FALSE;
ErrorIdValue := ComponentErrorNone;
StatusValue := BYTE#0;
END_METHOD

METHOD PUBLIC Snapshot : ComponentStatus
VAR
    Result : ComponentStatus;
END_VAR
Result.Ready := ReadyValue;
Result.Error := ErrorValue;
Result.ErrorId := ErrorIdValue;
Result.Status := StatusValue;
Snapshot := Result;
END_METHOD

METHOD PUBLIC SetLimits
VAR_INPUT
    Limits : RealRange;
END_VAR
IF Limits.High < Limits.Low THEN
    ErrorValue := TRUE;
    ErrorIdValue := ComponentErrorInvalidConfiguration;
    StatusValue := BYTE#1;
ELSE
    LowLimitValue := Limits.Low;
    HighLimitValue := Limits.High;
    ClearError();
END_IF;
END_METHOD

METHOD PUBLIC Update : BOOL
VAR_INPUT
    MeasuredValue : REAL;
END_VAR
IF NOT ReadyValue THEN
    ReadyValue := TRUE;
END_IF;
MeasuredValueValue := MeasuredValue;
IF MeasuredValueValue < LowLimitValue THEN
    QValue := FALSE;
    WindowValue := FALSE;
ELSIF MeasuredValueValue > HighLimitValue THEN
    QValue := TRUE;
    WindowValue := FALSE;
ELSE
    WindowValue := TRUE;
END_IF;
Update := QValue;
END_METHOD

PUBLIC PROPERTY Ready : BOOL
GET
    Ready := ReadyValue;
END_GET
END_PROPERTY

PUBLIC PROPERTY Error : BOOL
GET
    Error := ErrorValue;
END_GET
END_PROPERTY

PUBLIC PROPERTY ErrorId : WORD
GET
    ErrorId := ErrorIdValue;
END_GET
END_PROPERTY

PUBLIC PROPERTY Status : BYTE
GET
    Status := StatusValue;
END_GET
END_PROPERTY

PUBLIC PROPERTY MeasuredValue : REAL
GET
    MeasuredValue := MeasuredValueValue;
END_GET
END_PROPERTY

PUBLIC PROPERTY LowLimit : REAL
GET
    LowLimit := LowLimitValue;
END_GET
END_PROPERTY

PUBLIC PROPERTY HighLimit : REAL
GET
    HighLimit := HighLimitValue;
END_GET
END_PROPERTY

PUBLIC PROPERTY Q : BOOL
GET
    Q := QValue;
END_GET
END_PROPERTY

PUBLIC PROPERTY Window : BOOL
GET
    Window := WindowValue;
END_GET
END_PROPERTY
END_FUNCTION_BLOCK

FUNCTION_BLOCK TankLevelController IMPLEMENTS IComponent
VAR
    ReadyValue : BOOL;
    ErrorValue : BOOL;
    ErrorIdValue : WORD;
    StatusValue : BYTE;
    ValveValue : BOOL;
    AlarmValue : BOOL;
    MaxValveTimeValue : TIME;
    LevelDelayTimeValue : TIME;
    TankFb : TANK_LEVEL;
END_VAR

METHOD PUBLIC Initialize
ReadyValue := TRUE;
ClearError();
END_METHOD

METHOD PUBLIC Reset
TankFb(LEVEL := FALSE, LEAK := FALSE, ACLR := TRUE, MAX_VALVE_TIME := MaxValveTimeValue, LEVEL_DELAY_TIME := LevelDelayTimeValue);
ValveValue := TankFb.VALVE;
AlarmValue := TankFb.ALARM;
StatusValue := TankFb.STATUS;
ClearError();
END_METHOD

METHOD PUBLIC ClearError
ErrorValue := FALSE;
ErrorIdValue := ComponentErrorNone;
StatusValue := BYTE#0;
END_METHOD

METHOD PUBLIC Snapshot : ComponentStatus
VAR
    Result : ComponentStatus;
END_VAR
Result.Ready := ReadyValue;
Result.Error := ErrorValue;
Result.ErrorId := ErrorIdValue;
Result.Status := StatusValue;
Snapshot := Result;
END_METHOD

METHOD PUBLIC Configure
VAR_INPUT
    MaxValveTime : TIME;
    LevelDelayTime : TIME;
END_VAR
MaxValveTimeValue := MaxValveTime;
LevelDelayTimeValue := LevelDelayTime;
ClearError();
END_METHOD

METHOD PUBLIC Update : BOOL
VAR_INPUT
    LevelReached : BOOL;
    LeakDetected : BOOL;
    AlarmClear : BOOL;
END_VAR
TankFb(LEVEL := LevelReached, LEAK := LeakDetected, ACLR := AlarmClear, MAX_VALVE_TIME := MaxValveTimeValue, LEVEL_DELAY_TIME := LevelDelayTimeValue);
ValveValue := TankFb.VALVE;
AlarmValue := TankFb.ALARM;
StatusValue := TankFb.STATUS;
Update := ValveValue;
END_METHOD

PUBLIC PROPERTY Ready : BOOL
GET
    Ready := ReadyValue;
END_GET
END_PROPERTY

PUBLIC PROPERTY Error : BOOL
GET
    Error := ErrorValue;
END_GET
END_PROPERTY

PUBLIC PROPERTY ErrorId : WORD
GET
    ErrorId := ErrorIdValue;
END_GET
END_PROPERTY

PUBLIC PROPERTY Status : BYTE
GET
    Status := StatusValue;
END_GET
END_PROPERTY

PUBLIC PROPERTY Valve : BOOL
GET
    Valve := ValveValue;
END_GET
END_PROPERTY

PUBLIC PROPERTY Alarm : BOOL
GET
    Alarm := AlarmValue;
END_GET
END_PROPERTY
END_FUNCTION_BLOCK

FUNCTION_BLOCK HeatCurve IMPLEMENTS IComponent
VAR
    ReadyValue : BOOL;
    ErrorValue : BOOL;
    ErrorIdValue : WORD;
    StatusValue : BYTE;
    FlowTemperatureValue : REAL;
    HeatRequiredValue : BOOL;
    MaxFlowTemperatureValue : REAL := REAL#70.0;
    MinFlowTemperatureValue : REAL := REAL#25.0;
    ConfigFlowTemperatureValue : REAL := REAL#70.0;
    ConfigInsideTemperatureValue : REAL := REAL#20.0;
    ConfigOutsideTemperatureValue : REAL := REAL#-15.0;
    FlowDifferenceValue : REAL := REAL#10.0;
    CurveValue : REAL := REAL#1.33;
    HysteresisValue : REAL := REAL#3.0;
    HeatFb : HEAT_TEMP;
END_VAR

METHOD PUBLIC Initialize
ReadyValue := TRUE;
ClearError();
END_METHOD

METHOD PUBLIC Reset
FlowTemperatureValue := REAL#0.0;
HeatRequiredValue := FALSE;
ClearError();
END_METHOD

METHOD PUBLIC ClearError
ErrorValue := FALSE;
ErrorIdValue := ComponentErrorNone;
StatusValue := BYTE#0;
END_METHOD

METHOD PUBLIC Snapshot : ComponentStatus
VAR
    Result : ComponentStatus;
END_VAR
Result.Ready := ReadyValue;
Result.Error := ErrorValue;
Result.ErrorId := ErrorIdValue;
Result.Status := StatusValue;
Snapshot := Result;
END_METHOD

METHOD PUBLIC Configure
VAR_INPUT
    MaxFlowTemperature : REAL;
    MinFlowTemperature : REAL;
    ConfigFlowTemperature : REAL;
    ConfigInsideTemperature : REAL;
    ConfigOutsideTemperature : REAL;
    FlowDifference : REAL;
    Curve : REAL;
    Hysteresis : REAL;
END_VAR
MaxFlowTemperatureValue := MaxFlowTemperature;
MinFlowTemperatureValue := MinFlowTemperature;
ConfigFlowTemperatureValue := ConfigFlowTemperature;
ConfigInsideTemperatureValue := ConfigInsideTemperature;
ConfigOutsideTemperatureValue := ConfigOutsideTemperature;
FlowDifferenceValue := FlowDifference;
CurveValue := Curve;
HysteresisValue := Hysteresis;
ClearError();
END_METHOD

METHOD PUBLIC Update : REAL
VAR_INPUT
    OutsideTemperature : REAL;
    InsideTemperature : REAL;
    Offset : REAL;
    RequestedTemperature : REAL;
END_VAR
HeatFb(
    T_EXT := OutsideTemperature,
    T_INT := InsideTemperature,
    OFFSET := Offset,
    T_REQ := RequestedTemperature,
    TY_MAX := MaxFlowTemperatureValue,
    TY_MIN := MinFlowTemperatureValue,
    TY_CONFIG := ConfigFlowTemperatureValue,
    T_INT_CONFIG := ConfigInsideTemperatureValue,
    T_EXT_CONFIG := ConfigOutsideTemperatureValue,
    T_DIFF := FlowDifferenceValue,
    C := CurveValue,
    H := HysteresisValue
);
FlowTemperatureValue := HeatFb.TY;
HeatRequiredValue := HeatFb.HEAT;
Update := FlowTemperatureValue;
END_METHOD

PUBLIC PROPERTY Ready : BOOL
GET
    Ready := ReadyValue;
END_GET
END_PROPERTY

PUBLIC PROPERTY Error : BOOL
GET
    Error := ErrorValue;
END_GET
END_PROPERTY

PUBLIC PROPERTY ErrorId : WORD
GET
    ErrorId := ErrorIdValue;
END_GET
END_PROPERTY

PUBLIC PROPERTY Status : BYTE
GET
    Status := StatusValue;
END_GET
END_PROPERTY

PUBLIC PROPERTY FlowTemperature : REAL
GET
    FlowTemperature := FlowTemperatureValue;
END_GET
END_PROPERTY

PUBLIC PROPERTY HeatRequired : BOOL
GET
    HeatRequired := HeatRequiredValue;
END_GET
END_PROPERTY
END_FUNCTION_BLOCK

FUNCTION_BLOCK BoilerController IMPLEMENTS IComponent
VAR
    ReadyValue : BOOL;
    ErrorValue : BOOL;
    ErrorIdValue : WORD;
    StatusValue : BYTE;
    HeatValue : BOOL;
    BoilerErrorValue : BOOL;
    BoilerFb : BOILER;
END_VAR

METHOD PUBLIC Initialize
ReadyValue := TRUE;
ClearError();
END_METHOD

METHOD PUBLIC Reset
HeatValue := FALSE;
BoilerErrorValue := FALSE;
StatusValue := BYTE#0;
ClearError();
END_METHOD

METHOD PUBLIC ClearError
ErrorValue := FALSE;
ErrorIdValue := ComponentErrorNone;
StatusValue := BYTE#0;
END_METHOD

METHOD PUBLIC Snapshot : ComponentStatus
VAR
    Result : ComponentStatus;
END_VAR
Result.Ready := ReadyValue;
Result.Error := ErrorValue OR BoilerErrorValue;
Result.ErrorId := ErrorIdValue;
Result.Status := StatusValue;
Snapshot := Result;
END_METHOD

METHOD PUBLIC Update : BOOL
VAR_INPUT
    UpperTemperature : REAL;
    LowerTemperature : REAL;
    PressureOk : BOOL;
    Enabled : BOOL;
    Request1 : BOOL;
    Request2 : BOOL;
    Boost : BOOL;
END_VAR
BoilerFb(
    T_upper := UpperTemperature,
    T_lower := LowerTemperature,
    Pressure := PressureOk,
    enable := Enabled,
    Req_1 := Request1,
    Req_2 := Request2,
    Boost := Boost
);
HeatValue := BoilerFb.Heat;
BoilerErrorValue := BoilerFb.error;
StatusValue := BoilerFb.status;
Update := HeatValue;
END_METHOD

PUBLIC PROPERTY Ready : BOOL
GET
    Ready := ReadyValue;
END_GET
END_PROPERTY

PUBLIC PROPERTY Error : BOOL
GET
    Error := ErrorValue OR BoilerErrorValue;
END_GET
END_PROPERTY

PUBLIC PROPERTY ErrorId : WORD
GET
    ErrorId := ErrorIdValue;
END_GET
END_PROPERTY

PUBLIC PROPERTY Status : BYTE
GET
    Status := StatusValue;
END_GET
END_PROPERTY

PUBLIC PROPERTY Heat : BOOL
GET
    Heat := HeatValue;
END_GET
END_PROPERTY
END_FUNCTION_BLOCK

(* ---- device_drivers.st ---- *)
FUNCTION_BLOCK SingleOutputDriver IMPLEMENTS IComponent
VAR
    ReadyValue : BOOL;
    ErrorValue : BOOL;
    ErrorIdValue : WORD;
    StatusValue : BYTE;
    OutputValue : BOOL;
    ToggleModeValue : BOOL;
    TimeoutValue : TIME;
    DriverFb : DRIVER_1;
END_VAR

METHOD PUBLIC Initialize
ReadyValue := TRUE;
ClearError();
END_METHOD

METHOD PUBLIC Reset
DriverFb(SET_REQ := FALSE, IN := FALSE, RST := TRUE, Toggle_Mode := ToggleModeValue, Timeout := TimeoutValue);
OutputValue := DriverFb.Q;
ClearError();
END_METHOD

METHOD PUBLIC ClearError
ErrorValue := FALSE;
ErrorIdValue := ComponentErrorNone;
StatusValue := BYTE#0;
END_METHOD

METHOD PUBLIC Snapshot : ComponentStatus
VAR
    Result : ComponentStatus;
END_VAR
Result.Ready := ReadyValue;
Result.Error := ErrorValue;
Result.ErrorId := ErrorIdValue;
Result.Status := StatusValue;
Snapshot := Result;
END_METHOD

METHOD PUBLIC Configure
VAR_INPUT
    ToggleMode : BOOL;
    Timeout : TIME;
END_VAR
ToggleModeValue := ToggleMode;
TimeoutValue := Timeout;
ClearError();
END_METHOD

METHOD PUBLIC Update : BOOL
VAR_INPUT
    SetRequest : BOOL;
    Input : BOOL;
END_VAR
DriverFb(SET_REQ := SetRequest, IN := Input, RST := FALSE, Toggle_Mode := ToggleModeValue, Timeout := TimeoutValue);
OutputValue := DriverFb.Q;
Update := OutputValue;
END_METHOD

PUBLIC PROPERTY Ready : BOOL
GET
    Ready := ReadyValue;
END_GET
END_PROPERTY

PUBLIC PROPERTY Error : BOOL
GET
    Error := ErrorValue;
END_GET
END_PROPERTY

PUBLIC PROPERTY ErrorId : WORD
GET
    ErrorId := ErrorIdValue;
END_GET
END_PROPERTY

PUBLIC PROPERTY Status : BYTE
GET
    Status := StatusValue;
END_GET
END_PROPERTY

PUBLIC PROPERTY Output : BOOL
GET
    Output := OutputValue;
END_GET
END_PROPERTY
END_FUNCTION_BLOCK

(* ---- filters.st ---- *)
FUNCTION_BLOCK Pt1Filter IMPLEMENTS IPt1Filter
VAR
    ReadyValue : BOOL;
    ErrorValue : BOOL;
    ErrorIdValue : WORD;
    StatusValue : BYTE;
    OutputValue : REAL;
    TimeConstantValue : TIME := DefaultPt1TimeConstant;
    GainValue : REAL := DefaultPt1Gain;
    ResetRequested : BOOL;
    FilterFb : FT_PT1;
END_VAR

METHOD PUBLIC Initialize
ReadyValue := TRUE;
ClearError();
END_METHOD

METHOD PUBLIC Reset
ClearError();
OutputValue := REAL#0.0;
ResetRequested := TRUE;
END_METHOD

METHOD PUBLIC ClearError
ErrorValue := FALSE;
ErrorIdValue := ComponentErrorNone;
StatusValue := BYTE#0;
END_METHOD

METHOD PUBLIC Snapshot : ComponentStatus
VAR
    Result : ComponentStatus;
END_VAR
Result.Ready := ReadyValue;
Result.Error := ErrorValue;
Result.ErrorId := ErrorIdValue;
Result.Status := StatusValue;
Snapshot := Result;
END_METHOD

METHOD PUBLIC Configure
VAR_INPUT
    TimeConstant : TIME;
    Gain : REAL;
END_VAR
TimeConstantValue := TimeConstant;
GainValue := Gain;
ClearError();
END_METHOD

METHOD PUBLIC Update : REAL
VAR_INPUT
    Sample : REAL;
END_VAR
IF NOT ReadyValue THEN
    ReadyValue := TRUE;
END_IF;
IF ResetRequested THEN
    FilterFb(in := Sample, T := T#0s, K := GainValue);
    ResetRequested := FALSE;
ELSE
    FilterFb(in := Sample, T := TimeConstantValue, K := GainValue);
END_IF;
OutputValue := FilterFb.out;
Update := OutputValue;
END_METHOD

PUBLIC PROPERTY Ready : BOOL
GET
    Ready := ReadyValue;
END_GET
END_PROPERTY

PUBLIC PROPERTY Error : BOOL
GET
    Error := ErrorValue;
END_GET
END_PROPERTY

PUBLIC PROPERTY ErrorId : WORD
GET
    ErrorId := ErrorIdValue;
END_GET
END_PROPERTY

PUBLIC PROPERTY Status : BYTE
GET
    Status := StatusValue;
END_GET
END_PROPERTY

PUBLIC PROPERTY Output : REAL
GET
    Output := OutputValue;
END_GET
END_PROPERTY

PUBLIC PROPERTY TimeConstant : TIME
GET
    TimeConstant := TimeConstantValue;
END_GET
END_PROPERTY

PUBLIC PROPERTY Gain : REAL
GET
    Gain := GainValue;
END_GET
END_PROPERTY
END_FUNCTION_BLOCK

FUNCTION_BLOCK DerivativeFilter IMPLEMENTS IComponent
VAR
    ReadyValue : BOOL;
    ErrorValue : BOOL;
    ErrorIdValue : WORD;
    StatusValue : BYTE;
    OutputValue : REAL;
    GainValue : REAL := REAL#1.0;
    LastSample : REAL;
    LastTime : DWORD;
    Initialized : BOOL;
END_VAR

METHOD PUBLIC Initialize
ReadyValue := TRUE;
ClearError();
END_METHOD

METHOD PUBLIC Reset
Initialized := FALSE;
OutputValue := REAL#0.0;
ClearError();
END_METHOD

METHOD PUBLIC ClearError
ErrorValue := FALSE;
ErrorIdValue := ComponentErrorNone;
StatusValue := BYTE#0;
END_METHOD

METHOD PUBLIC Snapshot : ComponentStatus
VAR
    Result : ComponentStatus;
END_VAR
Result.Ready := ReadyValue;
Result.Error := ErrorValue;
Result.ErrorId := ErrorIdValue;
Result.Status := StatusValue;
Snapshot := Result;
END_METHOD

METHOD PUBLIC Configure
VAR_INPUT
    Gain : REAL;
END_VAR
GainValue := Gain;
ClearError();
END_METHOD

METHOD PUBLIC Update : REAL
VAR_INPUT
    Sample : REAL;
END_VAR
VAR
    NowTime : DWORD;
    DeltaUs : REAL;
END_VAR
NowTime := T_PLC_US();
DeltaUs := UDINT_TO_REAL(DWORD_TO_UDINT(NowTime) - DWORD_TO_UDINT(LastTime));
IF NOT Initialized THEN
    Initialized := TRUE;
    LastSample := Sample;
    OutputValue := REAL#0.0;
ELSIF DeltaUs > REAL#0.0 THEN
    OutputValue := (Sample - LastSample) / DeltaUs * REAL#1000000.0 * GainValue;
    LastSample := Sample;
ELSE
    OutputValue := REAL#0.0;
END_IF;
LastTime := NowTime;
Update := OutputValue;
END_METHOD

PUBLIC PROPERTY Ready : BOOL
GET
    Ready := ReadyValue;
END_GET
END_PROPERTY

PUBLIC PROPERTY Error : BOOL
GET
    Error := ErrorValue;
END_GET
END_PROPERTY

PUBLIC PROPERTY ErrorId : WORD
GET
    ErrorId := ErrorIdValue;
END_GET
END_PROPERTY

PUBLIC PROPERTY Status : BYTE
GET
    Status := StatusValue;
END_GET
END_PROPERTY

PUBLIC PROPERTY Output : REAL
GET
    Output := OutputValue;
END_GET
END_PROPERTY
END_FUNCTION_BLOCK

FUNCTION_BLOCK IntegratorFilter IMPLEMENTS IComponent
VAR
    ReadyValue : BOOL;
    ErrorValue : BOOL;
    ErrorIdValue : WORD;
    StatusValue : BYTE;
    OutputValue : REAL;
    LimitedValue : BOOL;
    GainValue : REAL := REAL#1.0;
    LowLimitValue : REAL := REAL#-1.0E37;
    HighLimitValue : REAL := REAL#1.0E37;
    ResetRequested : BOOL;
    FilterFb : FT_INT;
END_VAR

METHOD PUBLIC Initialize
ReadyValue := TRUE;
ClearError();
END_METHOD

METHOD PUBLIC Reset
ResetRequested := TRUE;
OutputValue := REAL#0.0;
LimitedValue := FALSE;
ClearError();
END_METHOD

METHOD PUBLIC ClearError
ErrorValue := FALSE;
ErrorIdValue := ComponentErrorNone;
StatusValue := BYTE#0;
END_METHOD

METHOD PUBLIC Snapshot : ComponentStatus
VAR
    Result : ComponentStatus;
END_VAR
Result.Ready := ReadyValue;
Result.Error := ErrorValue;
Result.ErrorId := ErrorIdValue;
Result.Status := StatusValue;
Snapshot := Result;
END_METHOD

METHOD PUBLIC Configure
VAR_INPUT
    Gain : REAL;
    Limits : RealRange;
END_VAR
IF Limits.High < Limits.Low THEN
    ErrorValue := TRUE;
    ErrorIdValue := ComponentErrorInvalidConfiguration;
    StatusValue := BYTE#1;
ELSE
    GainValue := Gain;
    LowLimitValue := Limits.Low;
    HighLimitValue := Limits.High;
    ClearError();
END_IF;
END_METHOD

METHOD PUBLIC Update : REAL
VAR_INPUT
    Sample : REAL;
    Run : BOOL;
END_VAR
FilterFb(IN := Sample, K := GainValue, RUN := Run, RST := ResetRequested, OUT_MIN := LowLimitValue, OUT_MAX := HighLimitValue);
ResetRequested := FALSE;
OutputValue := FilterFb.OUT;
LimitedValue := FilterFb.LIM;
Update := OutputValue;
END_METHOD

PUBLIC PROPERTY Ready : BOOL
GET
    Ready := ReadyValue;
END_GET
END_PROPERTY

PUBLIC PROPERTY Error : BOOL
GET
    Error := ErrorValue;
END_GET
END_PROPERTY

PUBLIC PROPERTY ErrorId : WORD
GET
    ErrorId := ErrorIdValue;
END_GET
END_PROPERTY

PUBLIC PROPERTY Status : BYTE
GET
    Status := StatusValue;
END_GET
END_PROPERTY

PUBLIC PROPERTY Output : REAL
GET
    Output := OutputValue;
END_GET
END_PROPERTY

PUBLIC PROPERTY Limited : BOOL
GET
    Limited := LimitedValue;
END_GET
END_PROPERTY
END_FUNCTION_BLOCK

FUNCTION_BLOCK Pt2Filter IMPLEMENTS IComponent
VAR
    ReadyValue : BOOL;
    ErrorValue : BOOL;
    ErrorIdValue : WORD;
    StatusValue : BYTE;
    OutputValue : REAL;
    TimeConstantValue : TIME := DefaultPt1TimeConstant;
    DampingValue : REAL := REAL#1.0;
    GainValue : REAL := DefaultPt1Gain;
    ResetRequested : BOOL;
    FilterFb : FT_PT2;
END_VAR

METHOD PUBLIC Initialize
ReadyValue := TRUE;
ClearError();
END_METHOD

METHOD PUBLIC Reset
ResetRequested := TRUE;
OutputValue := REAL#0.0;
ClearError();
END_METHOD

METHOD PUBLIC ClearError
ErrorValue := FALSE;
ErrorIdValue := ComponentErrorNone;
StatusValue := BYTE#0;
END_METHOD

METHOD PUBLIC Snapshot : ComponentStatus
VAR
    Result : ComponentStatus;
END_VAR
Result.Ready := ReadyValue;
Result.Error := ErrorValue;
Result.ErrorId := ErrorIdValue;
Result.Status := StatusValue;
Snapshot := Result;
END_METHOD

METHOD PUBLIC Configure
VAR_INPUT
    TimeConstant : TIME;
    Damping : REAL;
    Gain : REAL;
END_VAR
TimeConstantValue := TimeConstant;
DampingValue := Damping;
GainValue := Gain;
ClearError();
END_METHOD

METHOD PUBLIC Update : REAL
VAR_INPUT
    Sample : REAL;
END_VAR
IF ResetRequested THEN
    FilterFb(in := Sample, T := T#0s, D := DampingValue, K := GainValue);
    ResetRequested := FALSE;
ELSE
    FilterFb(in := Sample, T := TimeConstantValue, D := DampingValue, K := GainValue);
END_IF;
OutputValue := FilterFb.out;
Update := OutputValue;
END_METHOD

PUBLIC PROPERTY Ready : BOOL
GET
    Ready := ReadyValue;
END_GET
END_PROPERTY

PUBLIC PROPERTY Error : BOOL
GET
    Error := ErrorValue;
END_GET
END_PROPERTY

PUBLIC PROPERTY ErrorId : WORD
GET
    ErrorId := ErrorIdValue;
END_GET
END_PROPERTY

PUBLIC PROPERTY Status : BYTE
GET
    Status := StatusValue;
END_GET
END_PROPERTY

PUBLIC PROPERTY Output : REAL
GET
    Output := OutputValue;
END_GET
END_PROPERTY
END_FUNCTION_BLOCK

FUNCTION_BLOCK DelayLine16 IMPLEMENTS IComponent
VAR
    ReadyValue : BOOL;
    ErrorValue : BOOL;
    ErrorIdValue : WORD;
    StatusValue : BYTE;
    OutputValue : REAL;
    TriggeredValue : BOOL;
    DelayTimeValue : TIME := T#1s;
    DelayFb : FT_TN16;
END_VAR

METHOD PUBLIC Initialize
ReadyValue := TRUE;
ClearError();
END_METHOD

METHOD PUBLIC Reset
OutputValue := REAL#0.0;
TriggeredValue := FALSE;
ClearError();
END_METHOD

METHOD PUBLIC ClearError
ErrorValue := FALSE;
ErrorIdValue := ComponentErrorNone;
StatusValue := BYTE#0;
END_METHOD

METHOD PUBLIC Snapshot : ComponentStatus
VAR
    Result : ComponentStatus;
END_VAR
Result.Ready := ReadyValue;
Result.Error := ErrorValue;
Result.ErrorId := ErrorIdValue;
Result.Status := StatusValue;
Snapshot := Result;
END_METHOD

METHOD PUBLIC Configure
VAR_INPUT
    DelayTime : TIME;
END_VAR
DelayTimeValue := DelayTime;
ClearError();
END_METHOD

METHOD PUBLIC Update : REAL
VAR_INPUT
    Sample : REAL;
END_VAR
DelayFb(in := Sample, T := DelayTimeValue);
OutputValue := DelayFb.out;
TriggeredValue := DelayFb.trig;
Update := OutputValue;
END_METHOD

PUBLIC PROPERTY Ready : BOOL
GET
    Ready := ReadyValue;
END_GET
END_PROPERTY

PUBLIC PROPERTY Error : BOOL
GET
    Error := ErrorValue;
END_GET
END_PROPERTY

PUBLIC PROPERTY ErrorId : WORD
GET
    ErrorId := ErrorIdValue;
END_GET
END_PROPERTY

PUBLIC PROPERTY Status : BYTE
GET
    Status := StatusValue;
END_GET
END_PROPERTY

PUBLIC PROPERTY Output : REAL
GET
    Output := OutputValue;
END_GET
END_PROPERTY

PUBLIC PROPERTY Triggered : BOOL
GET
    Triggered := TriggeredValue;
END_GET
END_PROPERTY
END_FUNCTION_BLOCK

(* ---- generators.st ---- *)
FUNCTION_BLOCK PulseGenerator IMPLEMENTS IPulseGenerator
VAR
    ReadyValue : BOOL;
    ErrorValue : BOOL;
    ErrorIdValue : WORD;
    StatusValue : BYTE;
    EnabledValue : BOOL;
    OutputValue : BOOL;
    HighTimeValue : TIME := DefaultPulseHighTime;
    LowTimeValue : TIME := DefaultPulseLowTime;
    PulseFb : GEN_PULSE;
END_VAR

METHOD PUBLIC Initialize
ReadyValue := TRUE;
ClearError();
END_METHOD

METHOD PUBLIC Reset
EnabledValue := FALSE;
PulseFb(ENQ := FALSE, PTH := HighTimeValue, PTL := LowTimeValue);
OutputValue := PulseFb.Q;
ClearError();
END_METHOD

METHOD PUBLIC ClearError
ErrorValue := FALSE;
ErrorIdValue := ComponentErrorNone;
StatusValue := BYTE#0;
END_METHOD

METHOD PUBLIC Snapshot : ComponentStatus
VAR
    Result : ComponentStatus;
END_VAR
Result.Ready := ReadyValue;
Result.Error := ErrorValue;
Result.ErrorId := ErrorIdValue;
Result.Status := StatusValue;
Snapshot := Result;
END_METHOD

METHOD PUBLIC Configure
VAR_INPUT
    HighTime : TIME;
    LowTime : TIME;
END_VAR
HighTimeValue := HighTime;
LowTimeValue := LowTime;
ClearError();
END_METHOD

METHOD PUBLIC SetEnabled
VAR_INPUT
    Enabled : BOOL;
END_VAR
EnabledValue := Enabled;
ClearError();
END_METHOD

METHOD PUBLIC Update : BOOL
IF NOT ReadyValue THEN
    ReadyValue := TRUE;
END_IF;
PulseFb(ENQ := EnabledValue, PTH := HighTimeValue, PTL := LowTimeValue);
OutputValue := PulseFb.Q;
Update := OutputValue;
END_METHOD

PUBLIC PROPERTY Ready : BOOL
GET
    Ready := ReadyValue;
END_GET
END_PROPERTY

PUBLIC PROPERTY Error : BOOL
GET
    Error := ErrorValue;
END_GET
END_PROPERTY

PUBLIC PROPERTY ErrorId : WORD
GET
    ErrorId := ErrorIdValue;
END_GET
END_PROPERTY

PUBLIC PROPERTY Status : BYTE
GET
    Status := StatusValue;
END_GET
END_PROPERTY

PUBLIC PROPERTY Enabled : BOOL
GET
    Enabled := EnabledValue;
END_GET
END_PROPERTY

PUBLIC PROPERTY Output : BOOL
GET
    Output := OutputValue;
END_GET
END_PROPERTY

PUBLIC PROPERTY HighTime : TIME
GET
    HighTime := HighTimeValue;
END_GET
END_PROPERTY

PUBLIC PROPERTY LowTime : TIME
GET
    LowTime := LowTimeValue;
END_GET
END_PROPERTY
END_FUNCTION_BLOCK

FUNCTION_BLOCK RandomSignalGenerator IMPLEMENTS IComponent
VAR
    ReadyValue : BOOL;
    ErrorValue : BOOL;
    ErrorIdValue : WORD;
    StatusValue : BYTE;
    OutputValue : REAL;
    TriggeredValue : BOOL;
    PeriodValue : TIME := T#1s;
    AmplitudeValue : REAL := REAL#1.0;
    OffsetValue : REAL;
    GeneratorFb : GEN_RDM;
END_VAR

METHOD PUBLIC Initialize
ReadyValue := TRUE;
ClearError();
END_METHOD

METHOD PUBLIC Reset
OutputValue := REAL#0.0;
TriggeredValue := FALSE;
ClearError();
END_METHOD

METHOD PUBLIC ClearError
ErrorValue := FALSE;
ErrorIdValue := ComponentErrorNone;
StatusValue := BYTE#0;
END_METHOD

METHOD PUBLIC Snapshot : ComponentStatus
VAR
    Result : ComponentStatus;
END_VAR
Result.Ready := ReadyValue;
Result.Error := ErrorValue;
Result.ErrorId := ErrorIdValue;
Result.Status := StatusValue;
Snapshot := Result;
END_METHOD

METHOD PUBLIC Configure
VAR_INPUT
    Period : TIME;
    Amplitude : REAL;
    Offset : REAL;
END_VAR
PeriodValue := Period;
AmplitudeValue := Amplitude;
OffsetValue := Offset;
ClearError();
END_METHOD

METHOD PUBLIC Update : BOOL
GeneratorFb(PT := PeriodValue, AM := AmplitudeValue, OS := OffsetValue);
OutputValue := GeneratorFb.OUT;
TriggeredValue := GeneratorFb.Q;
Update := TriggeredValue;
END_METHOD

PUBLIC PROPERTY Ready : BOOL
GET
    Ready := ReadyValue;
END_GET
END_PROPERTY

PUBLIC PROPERTY Error : BOOL
GET
    Error := ErrorValue;
END_GET
END_PROPERTY

PUBLIC PROPERTY ErrorId : WORD
GET
    ErrorId := ErrorIdValue;
END_GET
END_PROPERTY

PUBLIC PROPERTY Status : BYTE
GET
    Status := StatusValue;
END_GET
END_PROPERTY

PUBLIC PROPERTY Output : REAL
GET
    Output := OutputValue;
END_GET
END_PROPERTY

PUBLIC PROPERTY Triggered : BOOL
GET
    Triggered := TriggeredValue;
END_GET
END_PROPERTY
END_FUNCTION_BLOCK

FUNCTION_BLOCK SineSignalGenerator IMPLEMENTS IComponent
VAR
    ReadyValue : BOOL;
    ErrorValue : BOOL;
    ErrorIdValue : WORD;
    StatusValue : BYTE;
    OutputValue : REAL;
    PositiveHalfValue : BOOL;
    PeriodValue : TIME := T#1s;
    AmplitudeValue : REAL := REAL#1.0;
    OffsetValue : REAL;
    DelayValue : REAL;
    GeneratorFb : GEN_SIN;
END_VAR

METHOD PUBLIC Initialize
ReadyValue := TRUE;
ClearError();
END_METHOD

METHOD PUBLIC Reset
OutputValue := REAL#0.0;
PositiveHalfValue := FALSE;
ClearError();
END_METHOD

METHOD PUBLIC ClearError
ErrorValue := FALSE;
ErrorIdValue := ComponentErrorNone;
StatusValue := BYTE#0;
END_METHOD

METHOD PUBLIC Snapshot : ComponentStatus
VAR
    Result : ComponentStatus;
END_VAR
Result.Ready := ReadyValue;
Result.Error := ErrorValue;
Result.ErrorId := ErrorIdValue;
Result.Status := StatusValue;
Snapshot := Result;
END_METHOD

METHOD PUBLIC Configure
VAR_INPUT
    Period : TIME;
    Amplitude : REAL;
    Offset : REAL;
    Delay : REAL;
END_VAR
PeriodValue := Period;
AmplitudeValue := Amplitude;
OffsetValue := Offset;
DelayValue := Delay;
ClearError();
END_METHOD

METHOD PUBLIC Update : REAL
GeneratorFb(PT := PeriodValue, AM := AmplitudeValue, OS := OffsetValue, DL := DelayValue);
OutputValue := GeneratorFb.OUT;
PositiveHalfValue := GeneratorFb.Q;
Update := OutputValue;
END_METHOD

PUBLIC PROPERTY Ready : BOOL
GET
    Ready := ReadyValue;
END_GET
END_PROPERTY

PUBLIC PROPERTY Error : BOOL
GET
    Error := ErrorValue;
END_GET
END_PROPERTY

PUBLIC PROPERTY ErrorId : WORD
GET
    ErrorId := ErrorIdValue;
END_GET
END_PROPERTY

PUBLIC PROPERTY Status : BYTE
GET
    Status := StatusValue;
END_GET
END_PROPERTY

PUBLIC PROPERTY Output : REAL
GET
    Output := OutputValue;
END_GET
END_PROPERTY

PUBLIC PROPERTY PositiveHalf : BOOL
GET
    PositiveHalf := PositiveHalfValue;
END_GET
END_PROPERTY
END_FUNCTION_BLOCK

FUNCTION_BLOCK SquareSignalGenerator IMPLEMENTS IComponent
VAR
    ReadyValue : BOOL;
    ErrorValue : BOOL;
    ErrorIdValue : WORD;
    StatusValue : BYTE;
    OutputValue : REAL;
    HighValue : BOOL;
    PeriodValue : TIME := T#1s;
    AmplitudeValue : REAL := REAL#1.0;
    OffsetValue : REAL;
    DutyCycleValue : REAL := REAL#0.5;
    DelayValue : REAL;
    GeneratorFb : GEN_SQR;
END_VAR

METHOD PUBLIC Initialize
ReadyValue := TRUE;
ClearError();
END_METHOD

METHOD PUBLIC Reset
OutputValue := REAL#0.0;
HighValue := FALSE;
ClearError();
END_METHOD

METHOD PUBLIC ClearError
ErrorValue := FALSE;
ErrorIdValue := ComponentErrorNone;
StatusValue := BYTE#0;
END_METHOD

METHOD PUBLIC Snapshot : ComponentStatus
VAR
    Result : ComponentStatus;
END_VAR
Result.Ready := ReadyValue;
Result.Error := ErrorValue;
Result.ErrorId := ErrorIdValue;
Result.Status := StatusValue;
Snapshot := Result;
END_METHOD

METHOD PUBLIC Configure
VAR_INPUT
    Period : TIME;
    Amplitude : REAL;
    Offset : REAL;
    DutyCycle : REAL;
    Delay : REAL;
END_VAR
PeriodValue := Period;
AmplitudeValue := Amplitude;
OffsetValue := Offset;
DutyCycleValue := DutyCycle;
DelayValue := Delay;
ClearError();
END_METHOD

METHOD PUBLIC Update : REAL
GeneratorFb(PT := PeriodValue, AM := AmplitudeValue, OS := OffsetValue, DC := DutyCycleValue, DL := DelayValue);
OutputValue := GeneratorFb.OUT;
HighValue := GeneratorFb.Q;
Update := OutputValue;
END_METHOD

PUBLIC PROPERTY Ready : BOOL
GET
    Ready := ReadyValue;
END_GET
END_PROPERTY

PUBLIC PROPERTY Error : BOOL
GET
    Error := ErrorValue;
END_GET
END_PROPERTY

PUBLIC PROPERTY ErrorId : WORD
GET
    ErrorId := ErrorIdValue;
END_GET
END_PROPERTY

PUBLIC PROPERTY Status : BYTE
GET
    Status := StatusValue;
END_GET
END_PROPERTY

PUBLIC PROPERTY Output : REAL
GET
    Output := OutputValue;
END_GET
END_PROPERTY

PUBLIC PROPERTY High : BOOL
GET
    High := HighValue;
END_GET
END_PROPERTY
END_FUNCTION_BLOCK

FUNCTION_BLOCK ByteRamp IMPLEMENTS IComponent
VAR
    ReadyValue : BOOL;
    ErrorValue : BOOL;
    ErrorIdValue : WORD;
    StatusValue : BYTE;
    OutputValue : BYTE;
    BusyValue : BOOL;
    HighValue : BOOL;
    LowValue : BOOL;
    RampFb : RMP_B;
END_VAR

METHOD PUBLIC Initialize
ReadyValue := TRUE;
ClearError();
END_METHOD

METHOD PUBLIC Reset
RampFb(SET_HIGH := FALSE, PT := T#0s, E := FALSE, UP := TRUE, RST := TRUE);
OutputValue := RampFb.OUT;
BusyValue := RampFb.BUSY;
HighValue := RampFb.HIGH;
LowValue := RampFb.LOW;
ClearError();
END_METHOD

METHOD PUBLIC ClearError
ErrorValue := FALSE;
ErrorIdValue := ComponentErrorNone;
StatusValue := BYTE#0;
END_METHOD

METHOD PUBLIC Snapshot : ComponentStatus
VAR
    Result : ComponentStatus;
END_VAR
Result.Ready := ReadyValue;
Result.Error := ErrorValue;
Result.ErrorId := ErrorIdValue;
Result.Status := StatusValue;
Snapshot := Result;
END_METHOD

METHOD PUBLIC Update : BYTE
VAR_INPUT
    SetHigh : BOOL;
    RampTime : TIME;
    Enabled : BOOL;
    Up : BOOL;
END_VAR
RampFb(SET_HIGH := SetHigh, PT := RampTime, E := Enabled, UP := Up, RST := FALSE);
OutputValue := RampFb.OUT;
BusyValue := RampFb.BUSY;
HighValue := RampFb.HIGH;
LowValue := RampFb.LOW;
Update := OutputValue;
END_METHOD

PUBLIC PROPERTY Ready : BOOL
GET
    Ready := ReadyValue;
END_GET
END_PROPERTY

PUBLIC PROPERTY Error : BOOL
GET
    Error := ErrorValue;
END_GET
END_PROPERTY

PUBLIC PROPERTY ErrorId : WORD
GET
    ErrorId := ErrorIdValue;
END_GET
END_PROPERTY

PUBLIC PROPERTY Status : BYTE
GET
    Status := StatusValue;
END_GET
END_PROPERTY

PUBLIC PROPERTY Output : BYTE
GET
    Output := OutputValue;
END_GET
END_PROPERTY

PUBLIC PROPERTY Busy : BOOL
GET
    Busy := BusyValue;
END_GET
END_PROPERTY
END_FUNCTION_BLOCK

FUNCTION_BLOCK WordRamp IMPLEMENTS IComponent
VAR
    ReadyValue : BOOL;
    ErrorValue : BOOL;
    ErrorIdValue : WORD;
    StatusValue : BYTE;
    OutputValue : WORD;
    BusyValue : BOOL;
    HighValue : BOOL;
    LowValue : BOOL;
    RampFb : RMP_W;
END_VAR

METHOD PUBLIC Initialize
ReadyValue := TRUE;
ClearError();
END_METHOD

METHOD PUBLIC Reset
RampFb(SET_HIGH := FALSE, PT := T#0s, E := FALSE, UP := TRUE, RST := TRUE);
OutputValue := RampFb.OUT;
BusyValue := RampFb.BUSY;
HighValue := RampFb.HIGH;
LowValue := RampFb.LOW;
ClearError();
END_METHOD

METHOD PUBLIC ClearError
ErrorValue := FALSE;
ErrorIdValue := ComponentErrorNone;
StatusValue := BYTE#0;
END_METHOD

METHOD PUBLIC Snapshot : ComponentStatus
VAR
    Result : ComponentStatus;
END_VAR
Result.Ready := ReadyValue;
Result.Error := ErrorValue;
Result.ErrorId := ErrorIdValue;
Result.Status := StatusValue;
Snapshot := Result;
END_METHOD

METHOD PUBLIC Update : WORD
VAR_INPUT
    SetHigh : BOOL;
    RampTime : TIME;
    Enabled : BOOL;
    Up : BOOL;
END_VAR
RampFb(SET_HIGH := SetHigh, PT := RampTime, E := Enabled, UP := Up, RST := FALSE);
OutputValue := RampFb.OUT;
BusyValue := RampFb.BUSY;
HighValue := RampFb.HIGH;
LowValue := RampFb.LOW;
Update := OutputValue;
END_METHOD

PUBLIC PROPERTY Ready : BOOL
GET
    Ready := ReadyValue;
END_GET
END_PROPERTY

PUBLIC PROPERTY Error : BOOL
GET
    Error := ErrorValue;
END_GET
END_PROPERTY

PUBLIC PROPERTY ErrorId : WORD
GET
    ErrorId := ErrorIdValue;
END_GET
END_PROPERTY

PUBLIC PROPERTY Status : BYTE
GET
    Status := StatusValue;
END_GET
END_PROPERTY

PUBLIC PROPERTY Output : WORD
GET
    Output := OutputValue;
END_GET
END_PROPERTY

PUBLIC PROPERTY Busy : BOOL
GET
    Busy := BusyValue;
END_GET
END_PROPERTY
END_FUNCTION_BLOCK

(* ---- logic.st ---- *)
FUNCTION_BLOCK Latch IMPLEMENTS IComponent
VAR
    ReadyValue : BOOL;
    ErrorValue : BOOL;
    ErrorIdValue : WORD;
    StatusValue : BYTE;
    OutputValue : BOOL;
    LatchFb : LTCH;
END_VAR

METHOD PUBLIC Initialize
ReadyValue := TRUE;
ClearError();
END_METHOD

METHOD PUBLIC Reset
LatchFb(DATA := FALSE, L := FALSE, RST := TRUE);
OutputValue := LatchFb.Q;
ClearError();
END_METHOD

METHOD PUBLIC ClearError
ErrorValue := FALSE;
ErrorIdValue := ComponentErrorNone;
StatusValue := BYTE#0;
END_METHOD

METHOD PUBLIC Snapshot : ComponentStatus
VAR
    Result : ComponentStatus;
END_VAR
Result.Ready := ReadyValue;
Result.Error := ErrorValue;
Result.ErrorId := ErrorIdValue;
Result.Status := StatusValue;
Snapshot := Result;
END_METHOD

METHOD PUBLIC Update : BOOL
VAR_INPUT
    Data : BOOL;
    Load : BOOL;
END_VAR
LatchFb(DATA := Data, L := Load, RST := FALSE);
OutputValue := LatchFb.Q;
Update := OutputValue;
END_METHOD

PUBLIC PROPERTY Ready : BOOL
GET
    Ready := ReadyValue;
END_GET
END_PROPERTY

PUBLIC PROPERTY Error : BOOL
GET
    Error := ErrorValue;
END_GET
END_PROPERTY

PUBLIC PROPERTY ErrorId : WORD
GET
    ErrorId := ErrorIdValue;
END_GET
END_PROPERTY

PUBLIC PROPERTY Status : BYTE
GET
    Status := StatusValue;
END_GET
END_PROPERTY

PUBLIC PROPERTY Output : BOOL
GET
    Output := OutputValue;
END_GET
END_PROPERTY
END_FUNCTION_BLOCK

FUNCTION_BLOCK ToggleSwitch IMPLEMENTS IComponent
VAR
    ReadyValue : BOOL;
    ErrorValue : BOOL;
    ErrorIdValue : WORD;
    StatusValue : BYTE;
    OutputValue : BOOL;
    ToggleFb : TOGGLE;
END_VAR

METHOD PUBLIC Initialize
ReadyValue := TRUE;
ClearError();
END_METHOD

METHOD PUBLIC Reset
ToggleFb(CLK := FALSE, RST := TRUE);
OutputValue := ToggleFb.Q;
ClearError();
END_METHOD

METHOD PUBLIC ClearError
ErrorValue := FALSE;
ErrorIdValue := ComponentErrorNone;
StatusValue := BYTE#0;
END_METHOD

METHOD PUBLIC Snapshot : ComponentStatus
VAR
    Result : ComponentStatus;
END_VAR
Result.Ready := ReadyValue;
Result.Error := ErrorValue;
Result.ErrorId := ErrorIdValue;
Result.Status := StatusValue;
Snapshot := Result;
END_METHOD

METHOD PUBLIC Update : BOOL
VAR_INPUT
    Clock : BOOL;
END_VAR
ToggleFb(CLK := Clock, RST := FALSE);
OutputValue := ToggleFb.Q;
Update := OutputValue;
END_METHOD

PUBLIC PROPERTY Ready : BOOL
GET
    Ready := ReadyValue;
END_GET
END_PROPERTY

PUBLIC PROPERTY Error : BOOL
GET
    Error := ErrorValue;
END_GET
END_PROPERTY

PUBLIC PROPERTY ErrorId : WORD
GET
    ErrorId := ErrorIdValue;
END_GET
END_PROPERTY

PUBLIC PROPERTY Status : BYTE
GET
    Status := StatusValue;
END_GET
END_PROPERTY

PUBLIC PROPERTY Output : BOOL
GET
    Output := OutputValue;
END_GET
END_PROPERTY
END_FUNCTION_BLOCK

FUNCTION_BLOCK DwordCounter IMPLEMENTS IComponent
VAR
    ReadyValue : BOOL;
    ErrorValue : BOOL;
    ErrorIdValue : WORD;
    StatusValue : BYTE;
    CountValue : DWORD;
    StepSizeValue : DWORD := DWORD#1;
    MaxValueValue : DWORD := DWORD#16#FFFFFFFF;
    CounterFb : COUNT_DR;
END_VAR

METHOD PUBLIC Initialize
ReadyValue := TRUE;
ClearError();
END_METHOD

METHOD PUBLIC Reset
CounterFb(SetIn := FALSE, IN := DWORD#0, UP := FALSE, DN := FALSE, StepSize := StepSizeValue, MX := MaxValueValue, RST := TRUE);
CountValue := CounterFb.CNT;
ClearError();
END_METHOD

METHOD PUBLIC ClearError
ErrorValue := FALSE;
ErrorIdValue := ComponentErrorNone;
StatusValue := BYTE#0;
END_METHOD

METHOD PUBLIC Snapshot : ComponentStatus
VAR
    Result : ComponentStatus;
END_VAR
Result.Ready := ReadyValue;
Result.Error := ErrorValue;
Result.ErrorId := ErrorIdValue;
Result.Status := StatusValue;
Snapshot := Result;
END_METHOD

METHOD PUBLIC Configure
VAR_INPUT
    StepSize : DWORD;
    MaxValue : DWORD;
END_VAR
StepSizeValue := StepSize;
MaxValueValue := MaxValue;
ClearError();
END_METHOD

METHOD PUBLIC SetValue
VAR_INPUT
    Value : DWORD;
END_VAR
CounterFb(SetIn := TRUE, IN := Value, UP := FALSE, DN := FALSE, StepSize := StepSizeValue, MX := MaxValueValue, RST := FALSE);
CountValue := CounterFb.CNT;
ClearError();
END_METHOD

METHOD PUBLIC Update : DWORD
VAR_INPUT
    Up : BOOL;
    Down : BOOL;
END_VAR
CounterFb(SetIn := FALSE, IN := DWORD#0, UP := Up, DN := Down, StepSize := StepSizeValue, MX := MaxValueValue, RST := FALSE);
CountValue := CounterFb.CNT;
Update := CountValue;
END_METHOD

PUBLIC PROPERTY Ready : BOOL
GET
    Ready := ReadyValue;
END_GET
END_PROPERTY

PUBLIC PROPERTY Error : BOOL
GET
    Error := ErrorValue;
END_GET
END_PROPERTY

PUBLIC PROPERTY ErrorId : WORD
GET
    ErrorId := ErrorIdValue;
END_GET
END_PROPERTY

PUBLIC PROPERTY Status : BYTE
GET
    Status := StatusValue;
END_GET
END_PROPERTY

PUBLIC PROPERTY Count : DWORD
GET
    Count := CountValue;
END_GET
END_PROPERTY
END_FUNCTION_BLOCK

FUNCTION_BLOCK ShiftRegister8 IMPLEMENTS IComponent
VAR
    ReadyValue : BOOL;
    ErrorValue : BOOL;
    ErrorIdValue : WORD;
    StatusValue : BYTE;
    OutputValue : BOOL;
    ShiftFb : SHR_8PLE;
END_VAR

METHOD PUBLIC Initialize
ReadyValue := TRUE;
ClearError();
END_METHOD

METHOD PUBLIC Reset
ShiftFb(Din := FALSE, Dload := BYTE#0, CLK := FALSE, UP := TRUE, LoadIn := FALSE, RST := TRUE);
OutputValue := ShiftFb.DOut;
ClearError();
END_METHOD

METHOD PUBLIC ClearError
ErrorValue := FALSE;
ErrorIdValue := ComponentErrorNone;
StatusValue := BYTE#0;
END_METHOD

METHOD PUBLIC Snapshot : ComponentStatus
VAR
    Result : ComponentStatus;
END_VAR
Result.Ready := ReadyValue;
Result.Error := ErrorValue;
Result.ErrorId := ErrorIdValue;
Result.Status := StatusValue;
Snapshot := Result;
END_METHOD

METHOD PUBLIC Update : BOOL
VAR_INPUT
    DataIn : BOOL;
    LoadValue : BYTE;
    Clock : BOOL;
    Up : BOOL;
    Load : BOOL;
END_VAR
ShiftFb(Din := DataIn, Dload := LoadValue, CLK := Clock, UP := Up, LoadIn := Load, RST := FALSE);
OutputValue := ShiftFb.DOut;
Update := OutputValue;
END_METHOD

PUBLIC PROPERTY Ready : BOOL
GET
    Ready := ReadyValue;
END_GET
END_PROPERTY

PUBLIC PROPERTY Error : BOOL
GET
    Error := ErrorValue;
END_GET
END_PROPERTY

PUBLIC PROPERTY ErrorId : WORD
GET
    ErrorId := ErrorIdValue;
END_GET
END_PROPERTY

PUBLIC PROPERTY Status : BYTE
GET
    Status := StatusValue;
END_GET
END_PROPERTY

PUBLIC PROPERTY Output : BOOL
GET
    Output := OutputValue;
END_GET
END_PROPERTY
END_FUNCTION_BLOCK

(* ---- measuring.st ---- *)
FUNCTION_BLOCK OntimeMeter IMPLEMENTS IComponent
VAR
    ReadyValue : BOOL;
    ErrorValue : BOOL;
    ErrorIdValue : WORD;
    StatusValue : BYTE;
    SecondsValue : UDINT;
    CyclesValue : UDINT;
    MeterFb : ONTIME;
END_VAR

METHOD PUBLIC Initialize
ReadyValue := TRUE;
ClearError();
END_METHOD

METHOD PUBLIC Reset
MeterFb(IN := FALSE, RST := TRUE, SECONDS := SecondsValue, CYCLES := CyclesValue);
ClearError();
END_METHOD

METHOD PUBLIC ClearError
ErrorValue := FALSE;
ErrorIdValue := ComponentErrorNone;
StatusValue := BYTE#0;
END_METHOD

METHOD PUBLIC Snapshot : ComponentStatus
VAR
    Result : ComponentStatus;
END_VAR
Result.Ready := ReadyValue;
Result.Error := ErrorValue;
Result.ErrorId := ErrorIdValue;
Result.Status := StatusValue;
Snapshot := Result;
END_METHOD

METHOD PUBLIC Update
VAR_INPUT
    Input : BOOL;
END_VAR
MeterFb(IN := Input, RST := FALSE, SECONDS := SecondsValue, CYCLES := CyclesValue);
END_METHOD

PUBLIC PROPERTY Ready : BOOL
GET
    Ready := ReadyValue;
END_GET
END_PROPERTY

PUBLIC PROPERTY Error : BOOL
GET
    Error := ErrorValue;
END_GET
END_PROPERTY

PUBLIC PROPERTY ErrorId : WORD
GET
    ErrorId := ErrorIdValue;
END_GET
END_PROPERTY

PUBLIC PROPERTY Status : BYTE
GET
    Status := StatusValue;
END_GET
END_PROPERTY

PUBLIC PROPERTY Seconds : UDINT
GET
    Seconds := SecondsValue;
END_GET
END_PROPERTY

PUBLIC PROPERTY Cycles : UDINT
GET
    Cycles := CyclesValue;
END_GET
END_PROPERTY
END_FUNCTION_BLOCK

FUNCTION_BLOCK CycleTimeMeter IMPLEMENTS IComponent
VAR
    ReadyValue : BOOL;
    ErrorValue : BOOL;
    ErrorIdValue : WORD;
    StatusValue : BYTE;
    MinValue : TIME;
    MaxValue : TIME;
    LastValue : TIME;
    SystemTimeValue : TIME;
    SystemDaysValue : INT;
    CyclesValue : DWORD;
    MeterFb : CYCLE_TIME;
END_VAR

METHOD PUBLIC Initialize
ReadyValue := TRUE;
ClearError();
END_METHOD

METHOD PUBLIC Reset
MeterFb(RST := TRUE);
MinValue := MeterFb.ct_min;
MaxValue := MeterFb.ct_max;
LastValue := MeterFb.ct_last;
SystemTimeValue := MeterFb.systime;
SystemDaysValue := MeterFb.sysdays;
CyclesValue := MeterFb.cycles;
ClearError();
END_METHOD

METHOD PUBLIC ClearError
ErrorValue := FALSE;
ErrorIdValue := ComponentErrorNone;
StatusValue := BYTE#0;
END_METHOD

METHOD PUBLIC Snapshot : ComponentStatus
VAR
    Result : ComponentStatus;
END_VAR
Result.Ready := ReadyValue;
Result.Error := ErrorValue;
Result.ErrorId := ErrorIdValue;
Result.Status := StatusValue;
Snapshot := Result;
END_METHOD

METHOD PUBLIC Update
VAR_INPUT
    ResetStatistics : BOOL;
END_VAR
MeterFb(RST := ResetStatistics);
MinValue := MeterFb.ct_min;
MaxValue := MeterFb.ct_max;
LastValue := MeterFb.ct_last;
SystemTimeValue := MeterFb.systime;
SystemDaysValue := MeterFb.sysdays;
CyclesValue := MeterFb.cycles;
END_METHOD

PUBLIC PROPERTY Ready : BOOL
GET
    Ready := ReadyValue;
END_GET
END_PROPERTY

PUBLIC PROPERTY Error : BOOL
GET
    Error := ErrorValue;
END_GET
END_PROPERTY

PUBLIC PROPERTY ErrorId : WORD
GET
    ErrorId := ErrorIdValue;
END_GET
END_PROPERTY

PUBLIC PROPERTY Status : BYTE
GET
    Status := StatusValue;
END_GET
END_PROPERTY

PUBLIC PROPERTY Cycles : DWORD
GET
    Cycles := CyclesValue;
END_GET
END_PROPERTY

PUBLIC PROPERTY LastCycleTime : TIME
GET
    LastCycleTime := LastValue;
END_GET
END_PROPERTY
END_FUNCTION_BLOCK

FUNCTION_BLOCK Calibrator IMPLEMENTS IComponent
VAR
    ReadyValue : BOOL;
    ErrorValue : BOOL;
    ErrorIdValue : WORD;
    StatusValue : BYTE;
    OutputValue : REAL;
    OffsetTargetValue : REAL;
    ScaleTargetValue : REAL := REAL#1.0;
    CalibratorFb : CALIBRATE;
END_VAR

METHOD PUBLIC Initialize
ReadyValue := TRUE;
ClearError();
END_METHOD

METHOD PUBLIC Reset
OutputValue := REAL#0.0;
ClearError();
END_METHOD

METHOD PUBLIC ClearError
ErrorValue := FALSE;
ErrorIdValue := ComponentErrorNone;
StatusValue := BYTE#0;
END_METHOD

METHOD PUBLIC Snapshot : ComponentStatus
VAR
    Result : ComponentStatus;
END_VAR
Result.Ready := ReadyValue;
Result.Error := ErrorValue;
Result.ErrorId := ErrorIdValue;
Result.Status := StatusValue;
Snapshot := Result;
END_METHOD

METHOD PUBLIC Configure
VAR_INPUT
    OffsetTarget : REAL;
    ScaleTarget : REAL;
END_VAR
OffsetTargetValue := OffsetTarget;
ScaleTargetValue := ScaleTarget;
ClearError();
END_METHOD

METHOD PUBLIC Update : REAL
VAR_INPUT
    Sample : REAL;
    CalibrateOffset : BOOL;
    CalibrateScale : BOOL;
END_VAR
CalibratorFb(X := Sample, CO := CalibrateOffset, CS := CalibrateScale, Y_Offset := OffsetTargetValue, Y_Scale := ScaleTargetValue);
OutputValue := CalibratorFb.Y;
Update := OutputValue;
END_METHOD

PUBLIC PROPERTY Ready : BOOL
GET
    Ready := ReadyValue;
END_GET
END_PROPERTY

PUBLIC PROPERTY Error : BOOL
GET
    Error := ErrorValue;
END_GET
END_PROPERTY

PUBLIC PROPERTY ErrorId : WORD
GET
    ErrorId := ErrorIdValue;
END_GET
END_PROPERTY

PUBLIC PROPERTY Status : BYTE
GET
    Status := StatusValue;
END_GET
END_PROPERTY

PUBLIC PROPERTY Output : REAL
GET
    Output := OutputValue;
END_GET
END_PROPERTY
END_FUNCTION_BLOCK

FUNCTION_BLOCK BarGraphMeter IMPLEMENTS IComponent
VAR
    ReadyValue : BOOL;
    ErrorValue : BOOL;
    ErrorIdValue : WORD;
    StatusValue : BYTE;
    LowValue : BOOL;
    Q1Value : BOOL;
    Q2Value : BOOL;
    Q3Value : BOOL;
    Q4Value : BOOL;
    Q5Value : BOOL;
    Q6Value : BOOL;
    HighValue : BOOL;
    AlarmValue : BOOL;
    TriggerLowValue : REAL;
    TriggerHighValue : REAL;
    AlarmLowValue : BOOL;
    AlarmHighValue : BOOL;
    LogScaleValue : BOOL;
    MeterFb : BAR_GRAPH;
END_VAR

METHOD PUBLIC Initialize
ReadyValue := TRUE;
ClearError();
END_METHOD

METHOD PUBLIC Reset
MeterFb(X := REAL#0.0, rst := TRUE, trigger_Low := TriggerLowValue, trigger_High := TriggerHighValue, Alarm_low := AlarmLowValue, Alarm_high := AlarmHighValue, log_scale := LogScaleValue);
CopyOutputs();
ClearError();
END_METHOD

METHOD PUBLIC ClearError
ErrorValue := FALSE;
ErrorIdValue := ComponentErrorNone;
StatusValue := BYTE#0;
END_METHOD

METHOD PUBLIC Snapshot : ComponentStatus
VAR
    Result : ComponentStatus;
END_VAR
Result.Ready := ReadyValue;
Result.Error := ErrorValue OR AlarmValue;
Result.ErrorId := ErrorIdValue;
Result.Status := StatusValue;
Snapshot := Result;
END_METHOD

METHOD PRIVATE CopyOutputs
LowValue := MeterFb.LOW;
Q1Value := MeterFb.Q1;
Q2Value := MeterFb.Q2;
Q3Value := MeterFb.Q3;
Q4Value := MeterFb.Q4;
Q5Value := MeterFb.Q5;
Q6Value := MeterFb.Q6;
HighValue := MeterFb.HIGH;
AlarmValue := MeterFb.Alarm;
StatusValue := MeterFb.Status;
END_METHOD

METHOD PUBLIC Configure
VAR_INPUT
    TriggerLow : REAL;
    TriggerHigh : REAL;
    AlarmLow : BOOL;
    AlarmHigh : BOOL;
    LogScale : BOOL;
END_VAR
TriggerLowValue := TriggerLow;
TriggerHighValue := TriggerHigh;
AlarmLowValue := AlarmLow;
AlarmHighValue := AlarmHigh;
LogScaleValue := LogScale;
ClearError();
END_METHOD

METHOD PUBLIC Update
VAR_INPUT
    Sample : REAL;
    ResetAlarm : BOOL;
END_VAR
MeterFb(X := Sample, rst := ResetAlarm, trigger_Low := TriggerLowValue, trigger_High := TriggerHighValue, Alarm_low := AlarmLowValue, Alarm_high := AlarmHighValue, log_scale := LogScaleValue);
CopyOutputs();
END_METHOD

PUBLIC PROPERTY Ready : BOOL
GET
    Ready := ReadyValue;
END_GET
END_PROPERTY

PUBLIC PROPERTY Error : BOOL
GET
    Error := ErrorValue OR AlarmValue;
END_GET
END_PROPERTY

PUBLIC PROPERTY ErrorId : WORD
GET
    ErrorId := ErrorIdValue;
END_GET
END_PROPERTY

PUBLIC PROPERTY Status : BYTE
GET
    Status := StatusValue;
END_GET
END_PROPERTY

PUBLIC PROPERTY Low : BOOL
GET
    Low := LowValue;
END_GET
END_PROPERTY

PUBLIC PROPERTY High : BOOL
GET
    High := HighValue;
END_GET
END_PROPERTY

PUBLIC PROPERTY Alarm : BOOL
GET
    Alarm := AlarmValue;
END_GET
END_PROPERTY
END_FUNCTION_BLOCK

(* ---- memory.st ---- *)
FUNCTION_BLOCK DwordFifo16 IMPLEMENTS IDwordQueue
VAR
    ReadyValue : BOOL;
    ErrorValue : BOOL;
    ErrorIdValue : WORD;
    StatusValue : BYTE;
    EmptyValue : BOOL := TRUE;
    FullValue : BOOL;
    ValueValue : DWORD;
    QueueFb : FIFO_16;
END_VAR

METHOD PUBLIC Initialize
ReadyValue := TRUE;
Reset();
END_METHOD

METHOD PUBLIC Reset
QueueFb(DIN := DWORD#0, E := TRUE, RD := FALSE, WD := FALSE, RST := TRUE);
ValueValue := QueueFb.DOUT;
EmptyValue := QueueFb.EMPTY;
FullValue := QueueFb.FULL;
ClearError();
END_METHOD

METHOD PUBLIC ClearError
ErrorValue := FALSE;
ErrorIdValue := ComponentErrorNone;
StatusValue := BYTE#0;
END_METHOD

METHOD PUBLIC Snapshot : ComponentStatus
VAR
    Result : ComponentStatus;
END_VAR
Result.Ready := ReadyValue;
Result.Error := ErrorValue;
Result.ErrorId := ErrorIdValue;
Result.Status := StatusValue;
Snapshot := Result;
END_METHOD

METHOD PUBLIC Push : BOOL
VAR_INPUT
    Value : DWORD;
END_VAR
IF FullValue THEN
    ErrorValue := TRUE;
    ErrorIdValue := ComponentErrorQueueFull;
    StatusValue := BYTE#1;
    Push := FALSE;
ELSE
    QueueFb(DIN := Value, E := TRUE, RD := FALSE, WD := TRUE, RST := FALSE);
    ValueValue := QueueFb.DOUT;
    EmptyValue := QueueFb.EMPTY;
    FullValue := QueueFb.FULL;
    Push := TRUE;
    ClearError();
END_IF;
END_METHOD

METHOD PUBLIC TryPop : BOOL
IF EmptyValue THEN
    TryPop := FALSE;
ELSE
    QueueFb(DIN := DWORD#0, E := TRUE, RD := TRUE, WD := FALSE, RST := FALSE);
    ValueValue := QueueFb.DOUT;
    EmptyValue := QueueFb.EMPTY;
    FullValue := QueueFb.FULL;
    TryPop := TRUE;
    ClearError();
END_IF;
END_METHOD

PUBLIC PROPERTY Ready : BOOL
GET
    Ready := ReadyValue;
END_GET
END_PROPERTY

PUBLIC PROPERTY Error : BOOL
GET
    Error := ErrorValue;
END_GET
END_PROPERTY

PUBLIC PROPERTY ErrorId : WORD
GET
    ErrorId := ErrorIdValue;
END_GET
END_PROPERTY

PUBLIC PROPERTY Status : BYTE
GET
    Status := StatusValue;
END_GET
END_PROPERTY

PUBLIC PROPERTY Empty : BOOL
GET
    Empty := EmptyValue;
END_GET
END_PROPERTY

PUBLIC PROPERTY Full : BOOL
GET
    Full := FullValue;
END_GET
END_PROPERTY

PUBLIC PROPERTY Value : DWORD
GET
    Value := ValueValue;
END_GET
END_PROPERTY

PUBLIC PROPERTY Capacity : UINT
GET
    Capacity := MaxDwordFifo16Capacity;
END_GET
END_PROPERTY
END_FUNCTION_BLOCK

FUNCTION_BLOCK DwordStack16 IMPLEMENTS IDwordStack
VAR
    ReadyValue : BOOL;
    ErrorValue : BOOL;
    ErrorIdValue : WORD;
    StatusValue : BYTE;
    EmptyValue : BOOL := TRUE;
    FullValue : BOOL;
    ValueValue : DWORD;
    StackFb : STACK_16;
END_VAR

METHOD PUBLIC Initialize
ReadyValue := TRUE;
Reset();
END_METHOD

METHOD PUBLIC Reset
StackFb(DIN := DWORD#0, E := TRUE, RD := FALSE, WD := FALSE, RST := TRUE);
ValueValue := StackFb.DOUT;
EmptyValue := StackFb.EMPTY;
FullValue := StackFb.FULL;
ClearError();
END_METHOD

METHOD PUBLIC ClearError
ErrorValue := FALSE;
ErrorIdValue := ComponentErrorNone;
StatusValue := BYTE#0;
END_METHOD

METHOD PUBLIC Snapshot : ComponentStatus
VAR
    Result : ComponentStatus;
END_VAR
Result.Ready := ReadyValue;
Result.Error := ErrorValue;
Result.ErrorId := ErrorIdValue;
Result.Status := StatusValue;
Snapshot := Result;
END_METHOD

METHOD PUBLIC Push : BOOL
VAR_INPUT
    Value : DWORD;
END_VAR
IF FullValue THEN
    ErrorValue := TRUE;
    ErrorIdValue := ComponentErrorQueueFull;
    StatusValue := BYTE#1;
    Push := FALSE;
ELSE
    StackFb(DIN := Value, E := TRUE, RD := FALSE, WD := TRUE, RST := FALSE);
    ValueValue := StackFb.DOUT;
    EmptyValue := StackFb.EMPTY;
    FullValue := StackFb.FULL;
    Push := TRUE;
    ClearError();
END_IF;
END_METHOD

METHOD PUBLIC TryPop : BOOL
IF EmptyValue THEN
    TryPop := FALSE;
ELSE
    StackFb(DIN := DWORD#0, E := TRUE, RD := TRUE, WD := FALSE, RST := FALSE);
    ValueValue := StackFb.DOUT;
    EmptyValue := StackFb.EMPTY;
    FullValue := StackFb.FULL;
    TryPop := TRUE;
    ClearError();
END_IF;
END_METHOD

PUBLIC PROPERTY Ready : BOOL
GET
    Ready := ReadyValue;
END_GET
END_PROPERTY

PUBLIC PROPERTY Error : BOOL
GET
    Error := ErrorValue;
END_GET
END_PROPERTY

PUBLIC PROPERTY ErrorId : WORD
GET
    ErrorId := ErrorIdValue;
END_GET
END_PROPERTY

PUBLIC PROPERTY Status : BYTE
GET
    Status := StatusValue;
END_GET
END_PROPERTY

PUBLIC PROPERTY Empty : BOOL
GET
    Empty := EmptyValue;
END_GET
END_PROPERTY

PUBLIC PROPERTY Full : BOOL
GET
    Full := FullValue;
END_GET
END_PROPERTY

PUBLIC PROPERTY Value : DWORD
GET
    Value := ValueValue;
END_GET
END_PROPERTY

PUBLIC PROPERTY Capacity : UINT
GET
    Capacity := MaxDwordStack16Capacity;
END_GET
END_PROPERTY
END_FUNCTION_BLOCK

FUNCTION_BLOCK DwordFifo32 IMPLEMENTS IDwordQueue
VAR
    ReadyValue : BOOL;
    ErrorValue : BOOL;
    ErrorIdValue : WORD;
    StatusValue : BYTE;
    EmptyValue : BOOL := TRUE;
    FullValue : BOOL;
    ValueValue : DWORD;
    QueueFb : FIFO_32;
END_VAR

METHOD PUBLIC Initialize
ReadyValue := TRUE;
Reset();
END_METHOD

METHOD PUBLIC Reset
QueueFb(DIN := DWORD#0, E := TRUE, RD := FALSE, WD := FALSE, RST := TRUE);
ValueValue := QueueFb.DOUT;
EmptyValue := QueueFb.EMPTY;
FullValue := QueueFb.FULL;
ClearError();
END_METHOD

METHOD PUBLIC ClearError
ErrorValue := FALSE;
ErrorIdValue := ComponentErrorNone;
StatusValue := BYTE#0;
END_METHOD

METHOD PUBLIC Snapshot : ComponentStatus
VAR
    Result : ComponentStatus;
END_VAR
Result.Ready := ReadyValue;
Result.Error := ErrorValue;
Result.ErrorId := ErrorIdValue;
Result.Status := StatusValue;
Snapshot := Result;
END_METHOD

METHOD PUBLIC Push : BOOL
VAR_INPUT
    Value : DWORD;
END_VAR
IF FullValue THEN
    ErrorValue := TRUE;
    ErrorIdValue := ComponentErrorQueueFull;
    StatusValue := BYTE#1;
    Push := FALSE;
ELSE
    QueueFb(DIN := Value, E := TRUE, RD := FALSE, WD := TRUE, RST := FALSE);
    ValueValue := QueueFb.DOUT;
    EmptyValue := QueueFb.EMPTY;
    FullValue := QueueFb.FULL;
    Push := TRUE;
    ClearError();
END_IF;
END_METHOD

METHOD PUBLIC TryPop : BOOL
IF EmptyValue THEN
    TryPop := FALSE;
ELSE
    QueueFb(DIN := DWORD#0, E := TRUE, RD := TRUE, WD := FALSE, RST := FALSE);
    ValueValue := QueueFb.DOUT;
    EmptyValue := QueueFb.EMPTY;
    FullValue := QueueFb.FULL;
    TryPop := TRUE;
    ClearError();
END_IF;
END_METHOD

PUBLIC PROPERTY Ready : BOOL
GET
    Ready := ReadyValue;
END_GET
END_PROPERTY

PUBLIC PROPERTY Error : BOOL
GET
    Error := ErrorValue;
END_GET
END_PROPERTY

PUBLIC PROPERTY ErrorId : WORD
GET
    ErrorId := ErrorIdValue;
END_GET
END_PROPERTY

PUBLIC PROPERTY Status : BYTE
GET
    Status := StatusValue;
END_GET
END_PROPERTY

PUBLIC PROPERTY Empty : BOOL
GET
    Empty := EmptyValue;
END_GET
END_PROPERTY

PUBLIC PROPERTY Full : BOOL
GET
    Full := FullValue;
END_GET
END_PROPERTY

PUBLIC PROPERTY Value : DWORD
GET
    Value := ValueValue;
END_GET
END_PROPERTY

PUBLIC PROPERTY Capacity : UINT
GET
    Capacity := MaxDwordFifo32Capacity;
END_GET
END_PROPERTY
END_FUNCTION_BLOCK

FUNCTION_BLOCK DwordStack32 IMPLEMENTS IDwordStack
VAR
    ReadyValue : BOOL;
    ErrorValue : BOOL;
    ErrorIdValue : WORD;
    StatusValue : BYTE;
    EmptyValue : BOOL := TRUE;
    FullValue : BOOL;
    ValueValue : DWORD;
    StackFb : STACK_32;
END_VAR

METHOD PUBLIC Initialize
ReadyValue := TRUE;
Reset();
END_METHOD

METHOD PUBLIC Reset
StackFb(DIN := DWORD#0, E := TRUE, RD := FALSE, WD := FALSE, RST := TRUE);
ValueValue := StackFb.DOUT;
EmptyValue := StackFb.EMPTY;
FullValue := StackFb.FULL;
ClearError();
END_METHOD

METHOD PUBLIC ClearError
ErrorValue := FALSE;
ErrorIdValue := ComponentErrorNone;
StatusValue := BYTE#0;
END_METHOD

METHOD PUBLIC Snapshot : ComponentStatus
VAR
    Result : ComponentStatus;
END_VAR
Result.Ready := ReadyValue;
Result.Error := ErrorValue;
Result.ErrorId := ErrorIdValue;
Result.Status := StatusValue;
Snapshot := Result;
END_METHOD

METHOD PUBLIC Push : BOOL
VAR_INPUT
    Value : DWORD;
END_VAR
IF FullValue THEN
    ErrorValue := TRUE;
    ErrorIdValue := ComponentErrorQueueFull;
    StatusValue := BYTE#1;
    Push := FALSE;
ELSE
    StackFb(DIN := Value, E := TRUE, RD := FALSE, WD := TRUE, RST := FALSE);
    ValueValue := StackFb.DOUT;
    EmptyValue := StackFb.EMPTY;
    FullValue := StackFb.FULL;
    Push := TRUE;
    ClearError();
END_IF;
END_METHOD

METHOD PUBLIC TryPop : BOOL
IF EmptyValue THEN
    TryPop := FALSE;
ELSE
    StackFb(DIN := DWORD#0, E := TRUE, RD := TRUE, WD := FALSE, RST := FALSE);
    ValueValue := StackFb.DOUT;
    EmptyValue := StackFb.EMPTY;
    FullValue := StackFb.FULL;
    TryPop := TRUE;
    ClearError();
END_IF;
END_METHOD

PUBLIC PROPERTY Ready : BOOL
GET
    Ready := ReadyValue;
END_GET
END_PROPERTY

PUBLIC PROPERTY Error : BOOL
GET
    Error := ErrorValue;
END_GET
END_PROPERTY

PUBLIC PROPERTY ErrorId : WORD
GET
    ErrorId := ErrorIdValue;
END_GET
END_PROPERTY

PUBLIC PROPERTY Status : BYTE
GET
    Status := StatusValue;
END_GET
END_PROPERTY

PUBLIC PROPERTY Empty : BOOL
GET
    Empty := EmptyValue;
END_GET
END_PROPERTY

PUBLIC PROPERTY Full : BOOL
GET
    Full := FullValue;
END_GET
END_PROPERTY

PUBLIC PROPERTY Value : DWORD
GET
    Value := ValueValue;
END_GET
END_PROPERTY

PUBLIC PROPERTY Capacity : UINT
GET
    Capacity := MaxDwordStack32Capacity;
END_GET
END_PROPERTY
END_FUNCTION_BLOCK

(* ---- unit_converter.st ---- *)
FUNCTION_BLOCK UnitConverter IMPLEMENTS IUnitConverter
VAR
    ReadyValue : BOOL;
    ErrorValue : BOOL;
    ErrorIdValue : WORD;
    StatusValue : BYTE;
    EnergyFb : ENERGY;
END_VAR

METHOD PUBLIC Initialize
ReadyValue := TRUE;
ClearError();
END_METHOD

METHOD PUBLIC Reset
ClearError();
END_METHOD

METHOD PUBLIC ClearError
ErrorValue := FALSE;
ErrorIdValue := ComponentErrorNone;
StatusValue := BYTE#0;
END_METHOD

METHOD PUBLIC Snapshot : ComponentStatus
VAR
    Result : ComponentStatus;
END_VAR
Result.Ready := ReadyValue;
Result.Error := ErrorValue;
Result.ErrorId := ErrorIdValue;
Result.Status := StatusValue;
Snapshot := Result;
END_METHOD

METHOD PUBLIC KelvinFromCelsius : REAL
VAR_INPUT
    Celsius : REAL;
END_VAR
OSCAT_BASIC_Constants();
KelvinFromCelsius := C_TO_K(Celsius := Celsius);
END_METHOD

METHOD PUBLIC FahrenheitFromCelsius : REAL
VAR_INPUT
    Celsius : REAL;
END_VAR
FahrenheitFromCelsius := C_TO_F(celsius := Celsius);
END_METHOD

METHOD PUBLIC CelsiusFromKelvin : REAL
VAR_INPUT
    Kelvin : REAL;
END_VAR
OSCAT_BASIC_Constants();
CelsiusFromKelvin := K_TO_C(Kelvin := Kelvin);
END_METHOD

METHOD PUBLIC CelsiusFromFahrenheit : REAL
VAR_INPUT
    Fahrenheit : REAL;
END_VAR
OSCAT_BASIC_Constants();
CelsiusFromFahrenheit := F_TO_C(fahrenheit := Fahrenheit);
END_METHOD

METHOD PUBLIC MetersPerSecondFromKilometersPerHour : REAL
VAR_INPUT
    Kmh : REAL;
END_VAR
MetersPerSecondFromKilometersPerHour := KMH_TO_MS(kmh := Kmh);
END_METHOD

METHOD PUBLIC KilometersPerHourFromMetersPerSecond : REAL
VAR_INPUT
    Mps : REAL;
END_VAR
KilometersPerHourFromMetersPerSecond := MS_TO_KMH(ms := Mps);
END_METHOD

METHOD PUBLIC BeaufortFromMetersPerSecond : INT
VAR_INPUT
    Mps : REAL;
END_VAR
BeaufortFromMetersPerSecond := MS_TO_BFT(MS := Mps);
END_METHOD

METHOD PUBLIC AngularFrequencyFromHertz : REAL
VAR_INPUT
    Frequency : REAL;
END_VAR
OSCAT_BASIC_Constants();
AngularFrequencyFromHertz := F_TO_OM(F := Frequency);
END_METHOD

METHOD PUBLIC HertzFromAngularFrequency : REAL
VAR_INPUT
    AngularFrequency : REAL;
END_VAR
OSCAT_BASIC_Constants();
HertzFromAngularFrequency := OM_TO_F(OM := AngularFrequency);
END_METHOD

METHOD PUBLIC PeriodFromHertz : TIME
VAR_INPUT
    Frequency : REAL;
END_VAR
PeriodFromHertz := F_TO_PT(F := Frequency);
END_METHOD

METHOD PUBLIC HertzFromPeriod : REAL
VAR_INPUT
    Period : TIME;
END_VAR
HertzFromPeriod := PT_TO_F(PT := Period);
END_METHOD

METHOD PUBLIC WattHoursFromJoules : REAL
VAR_INPUT
    Joule : REAL;
END_VAR
EnergyFb(J := Joule, C := REAL#0.0, Wh := REAL#0.0);
WattHoursFromJoules := EnergyFb.YWh;
END_METHOD

METHOD PUBLIC JoulesFromWattHours : REAL
VAR_INPUT
    WattHour : REAL;
END_VAR
EnergyFb(J := REAL#0.0, C := REAL#0.0, Wh := WattHour);
JoulesFromWattHours := EnergyFb.YJ;
END_METHOD

METHOD PUBLIC JoulesFromCalories : REAL
VAR_INPUT
    Calorie : REAL;
END_VAR
EnergyFb(J := REAL#0.0, C := Calorie, Wh := REAL#0.0);
JoulesFromCalories := EnergyFb.YJ;
END_METHOD

METHOD PUBLIC CaloriesFromJoules : REAL
VAR_INPUT
    Joule : REAL;
END_VAR
EnergyFb(J := Joule, C := REAL#0.0, Wh := REAL#0.0);
CaloriesFromJoules := EnergyFb.YC;
END_METHOD

PUBLIC PROPERTY Ready : BOOL
GET
    Ready := ReadyValue;
END_GET
END_PROPERTY

PUBLIC PROPERTY Error : BOOL
GET
    Error := ErrorValue;
END_GET
END_PROPERTY

PUBLIC PROPERTY ErrorId : WORD
GET
    ErrorId := ErrorIdValue;
END_GET
END_PROPERTY

PUBLIC PROPERTY Status : BYTE
GET
    Status := StatusValue;
END_GET
END_PROPERTY
END_FUNCTION_BLOCK
